// TwinCAT 3 PLC project Intecre_TwinSafeModels
// Title: Intecre.TwinSAFE.Models
// Company: Intecre Ltd
// Author: Mark Lazarides
// ProjectVersion: 0.5.0.3
// Description: Functional models of the TwinSAFE logic function blocks and TwinSAFE group, for trialling safety applications and their interaction with the standard PLC. 0.4.2.0 - T_SafeFunctionBlockBase sets State to Run / Stop before Process; user FBs need no State logic. 0.4.1.0 - corrects call issue with Example_UserFBs 0.4.0.0 - Adds the eight channel (EL1918) and two channel (EL2912) terminal models. 0.3.0.0 - Adds User FB examples, demonstrating extension.
// ProgramVersion: 3.1.4026.25
// libraries:
//   Intecre.Utilities, * (Intecre Ltd)
//   Tc2_Standard, * (Beckhoff Automation GmbH)
//   Tc2_System, * (Beckhoff Automation GmbH)
//   Tc3_Module, * (Beckhoff Automation GmbH)
//   TcUnit, * (www.tcunit.org)
// project tree:
//   / PlcTask.TcTTO
//   Core/ F_NormaliseSafeInput.TcPOU, F_SafeResetTimeOk.TcPOU, F_SafeInputValue.TcPOU, T_SafeConnection.TcPOU, T_SafeFunctionBlockBase.TcPOU, T_SafeGroup.TcPOU, T_SafeInputPair.TcPOU, T_SafeInputTerminal.TcPOU, T_SafeInputTerminal8.TcPOU, T_SafeOutputTerminal.TcPOU, T_SafeOutputTerminal2.TcPOU
//   DUTs/ E_SafeConnectionError.TcDUT, E_SafeConnectionState.TcDUT, E_SafeEdmState.TcDUT, E_SafeFbState.TcDUT, E_SafeGroupDiag.TcDUT, E_SafeGroupState.TcDUT, E_SafeLatchState.TcDUT, E_SafeMonState.TcDUT, E_SafeMutingState.TcDUT, E_SafeTonState.TcDUT, E_SafeTwoHandState.TcDUT, ST_SafeConnShutdownParameters.TcDUT, ST_SafeEStopParameters.TcDUT, ST_SafeEdmParameters.TcDUT, ST_SafeLatchParameters.TcDUT, ST_SafeLogicParameters.TcDUT, ST_SafeMonParameters.TcDUT, ST_SafeMutingParameters.TcDUT, ST_SafeOpModeParameters.TcDUT, ST_SafeTimerParameters.TcDUT, ST_SafeTwoHandParameters.TcDUT
//   Examples/Example_UserFbs/ T_SafePulse_UserFB.TcPOU, T_SafeRTrig_UserFB.TcPOU
//   Examples/ PRG_EStopExample.TcPOU, PRG_EStopExample_CFC.TcPOU
//   FunctionBlocks/ T_SafeAnd.TcPOU, T_SafeConnShutdown.TcPOU, T_SafeDecouple.TcPOU, T_SafeEStop.TcPOU, T_SafeEdm.TcPOU, T_SafeMon.TcPOU, T_SafeMuting.TcPOU, T_SafeOpMode.TcPOU, T_SafeOr.TcPOU, T_SafeRs.TcPOU, T_SafeSr.TcPOU, T_SafeTof.TcPOU, T_SafeTon.TcPOU, T_SafeTwoHand.TcPOU, T_SafeXor.TcPOU
//   Params/ SafeModelParams.TcGVL
//   Project Information/ F_GetCompany.TcPOU, F_GetTitle.TcPOU, F_GetVersion.TcPOU
//   Tests/ T_SafeCfcTestSuite.TcPOU, PRG_TestRunner.TcPOU, T_SafeAnd_Tests.TcPOU, T_SafeAnd_Tests_CFC.TcPOU, T_SafeConnShutdown_Tests.TcPOU, T_SafeConnShutdown_Tests_CFC.TcPOU, T_SafeConnection_Tests.TcPOU, T_SafeConnection_Tests_CFC.TcPOU, T_SafeDecouple_Tests.TcPOU, T_SafeDecouple_Tests_CFC.TcPOU, T_SafeEStop_Tests.TcPOU, T_SafeEStop_Tests_CFC.TcPOU, T_SafeEdm_Tests.TcPOU, T_SafeEdm_Tests_CFC.TcPOU, T_SafeGroup_Tests.TcPOU, T_SafeGroup_Tests_CFC.TcPOU, T_SafeInputPair_Tests.TcPOU, T_SafeInputPair_Tests_CFC.TcPOU, T_SafeInputTerminal8_Tests.TcPOU, T_SafeMon_Tests.TcPOU, T_SafeMon_Tests_CFC.TcPOU, T_SafeMuting_Tests.TcPOU, T_SafeMuting_Tests_CFC.TcPOU, T_SafeOpMode_Tests.TcPOU, T_SafeOpMode_Tests_CFC.TcPOU, T_SafeOr_Tests.TcPOU, T_SafeOr_Tests_CFC.TcPOU, T_SafeOutputTerminal2_Tests.TcPOU, T_SafeRs_Tests.TcPOU, T_SafeRs_Tests_CFC.TcPOU, T_SafeSr_Tests.TcPOU, T_SafeSr_Tests_CFC.TcPOU, T_SafeTof_Tests.TcPOU, T_SafeTof_Tests_CFC.TcPOU, T_SafeTon_Tests.TcPOU, T_SafeTon_Tests_CFC.TcPOU, T_SafeTwoHand_Tests.TcPOU, T_SafeTwoHand_Tests_CFC.TcPOU, T_SafeXor_Tests.TcPOU, T_SafeXor_Tests_CFC.TcPOU
//   Tests/User_FB_Tests/ T_SafePulse_UserFB_Tests.TcPOU, T_SafePulse_UserFB_Tests_CFC.TcPOU, T_SafeRTrig_UserFB_Tests.TcPOU, T_SafeRTrig_UserFB_Tests_CFC.TcPOU
//   Version/ Global_Version.TcGVL
// real-time tasks:
//   TASK PlcTask: cycle T#10ms, priority 20, ADS port 350

CONFIGURATION Intecre_TwinSafeModels
    RESOURCE PLC ON TwinCAT3
        TASK PlcTask(INTERVAL := T#10ms, PRIORITY := 20);
        PROGRAM PRG_TestRunner WITH PlcTask : PRG_TestRunner;
        PROGRAM PRG_EStopExample WITH PlcTask : PRG_EStopExample;
        PROGRAM PRG_EStopExample_CFC WITH PlcTask : PRG_EStopExample_CFC;
    END_RESOURCE
END_CONFIGURATION

// ---- DUTs/E_SafeConnectionError.TcDUT
// TwinSAFE connection error codes (low nibble of the connection Diag byte).
{attribute 'qualified_only'}
{attribute 'to_string'}
TYPE
E_SafeConnectionError :
(
    NoError := 0,
    InvalidCommand := 1,
    UnknownCommand := 2,
    InvalidConnectionId := 3,
    InvalidCrc := 4,
    WatchdogElapsed := 5,
    InvalidFsoeAddress := 6,
    InvalidData := 7,
    InvalidComParameterLength := 8,
    InvalidComParameters := 9,
    InvalidUserParameterLength := 10,
    InvalidUserParameters := 11,
    FsoeMasterReset := 12,
    SlaveModuleError := 13,
    OutputModuleError := 14,
    SlaveNotStarted := 15
) BYTE;
END_TYPE

// ---- DUTs/E_SafeConnectionState.TcDUT
// TwinSAFE (FSoE) connection state codes.
{attribute 'qualified_only'}
{attribute 'to_string'}
TYPE
E_SafeConnectionState :
(
    Reset := 100,
    Session := 101,
    Connection := 102,
    Parameter := 103,
    Data := 104,
    Shutdown := 105,
    ShutdownDeactive := 106
) BYTE;
END_TYPE

// ---- DUTs/E_SafeEdmState.TcDUT
// FB EDM state codes.
{attribute 'qualified_only'}
{attribute 'to_string'}
TYPE
E_SafeEdmState :
(
    Undefined := 0,
    Stop := 2,
    Error := 4,
    Reset := 5,
    MonOff := 14,
    MonOn := 15
) BYTE;
END_TYPE

// ---- DUTs/E_SafeFbState.TcDUT
// TwinSAFE function block state codes shared by most FBs (Map State value).
// Error is also the state of a block whose configuration the TwinSAFE Safety Editor refuses (too few
// inputs connected, a required input unwired, an invalid EDM reset time): the block then sets Error,
// diagnostic bit 15 (16#8000), which no TwinSAFE FB uses, and stays in Error through every ErrAck.
// See T_SafeFunctionBlockBase.
{attribute 'qualified_only'}
{attribute 'to_string'}
TYPE
E_SafeFbState :
(
    Undefined := 0,
    Run := 1,
    Stop := 2,
    Safe := 3,
    Error := 4,
    Reset := 5,
    Start := 6,
    ErrorDelay := 7,
    DelayOut := 8
) BYTE;
END_TYPE

// ---- DUTs/E_SafeGroupDiag.TcDUT
// TwinSAFE group diagnostic codes (EL/EJ6910).
{attribute 'qualified_only'}
{attribute 'to_string'}
TYPE
E_SafeGroupDiag :
(
    NoError := 0,
    FbError := 1,
    ComError := 2,
    ModuleError := 3,
    CmpError := 4,
    DeactivateError := 5,
    RestartError := 6
) BYTE;
END_TYPE

// ---- DUTs/E_SafeGroupState.TcDUT
// TwinSAFE group state codes (EL/EJ6910).
{attribute 'qualified_only'}
{attribute 'to_string'}
TYPE
E_SafeGroupState :
(
    Undefined := 0,
    Run := 1,
    Stop := 2,
    Safe := 3,
    Error := 4,
    Reset := 5,
    Start := 6,
    StopError := 7,
    Deactive := 16,
    WaitComError := 17
) BYTE;
END_TYPE

// ---- DUTs/E_SafeLatchState.TcDUT
// FB RS and FB SR state codes.
{attribute 'qualified_only'}
{attribute 'to_string'}
TYPE
E_SafeLatchState :
(
    Undefined := 0,
    Stop := 2,
    Safe := 3,
    Set := 9
) BYTE;
END_TYPE

// ---- DUTs/E_SafeMonState.TcDUT
// FB MON state codes.
{attribute 'qualified_only'}
{attribute 'to_string'}
TYPE
E_SafeMonState :
(
    Undefined := 0,
    Run := 1,
    Stop := 2,
    Safe := 3,
    Error := 4,
    Reset := 5,
    Start := 6,
    ErrorDelay := 7,
    DelayOut := 8,
    FuncTest := 9
) BYTE;
END_TYPE

// ---- DUTs/E_SafeMutingState.TcDUT
// FB MUTING state codes.
{attribute 'qualified_only'}
{attribute 'to_string'}
TYPE
E_SafeMutingState :
(
    Undefined := 0,
    Run := 1,
    Stop := 2,
    Safe := 3,
    Error := 4,
    Reset := 5,
    DelayOut := 8,
    Muting1 := 9,
    Muting2 := 10,
    Muting3 := 11,
    Muting4 := 12,
    Muting5 := 13,
    Muting6 := 14,
    Muting7 := 15,
    Muting8 := 16,
    Muting9 := 17
) BYTE;
END_TYPE

// ---- DUTs/E_SafeTonState.TcDUT
// FB TON state codes.
{attribute 'qualified_only'}
{attribute 'to_string'}
TYPE
E_SafeTonState :
(
    Undefined := 0,
    Run := 1,
    Stop := 2,
    Safe := 3,
    DelayIn := 9
) BYTE;
END_TYPE

// ---- DUTs/E_SafeTwoHandState.TcDUT
// FB TWOHAND state codes.
{attribute 'qualified_only'}
{attribute 'to_string'}
TYPE
E_SafeTwoHandState :
(
    Undefined := 0,
    Run := 1,
    Stop := 2,
    Safe := 3,
    Error := 4,
    Reset := 5,
    OneButton := 11,
    TwoButton := 12,
    Release := 13
) BYTE;
END_TYPE

// ---- DUTs/ST_SafeConnShutdownParameters.TcDUT
// Parameters of FB CONNECTION SHUTDOWN.
TYPE
ST_SafeConnShutdownParameters :
STRUCT
    Deactivate1MakeContact : BOOL;
    Deactivate2MakeContact : BOOL;
    DiscrepancyTime : TIME;
    SafeInputsAfterDiscError : BOOL; // Safety Editor checkbox 'Safe Inputs after Disc Error', FALSE for a new block:
        // TRUE makes both channels of the pair that raised a discrepancy error return to the safe state together
        // before ErrAck can clear it
END_STRUCT
END_TYPE

// ---- DUTs/ST_SafeEStopParameters.TcDUT
// Parameters of FB ESTOP (port and FB properties of the Safety Editor).
// Ports are active when connected; a pair is two channel when both ports are connected.
TYPE
ST_SafeEStopParameters :
STRUCT
    EStopIn1MakeContact : BOOL; // FALSE = break contact (0 requests the safe state); TRUE = make contact
    EStopIn2MakeContact : BOOL;
    EStopIn3MakeContact : BOOL;
    EStopIn4MakeContact : BOOL;
    EStopIn5MakeContact : BOOL;
    EStopIn6MakeContact : BOOL;
    EStopIn7MakeContact : BOOL;
    EStopIn8MakeContact : BOOL;
    DiscrepancyTime1 : TIME; // EStopIn1 / EStopIn2. T#0S = no discrepancy monitoring
    DiscrepancyTime2 : TIME; // EStopIn3 / EStopIn4
    DiscrepancyTime3 : TIME; // EStopIn5 / EStopIn6
    DiscrepancyTime4 : TIME; // EStopIn7 / EStopIn8
    DelayTime : TIME; // switch-off delay of EStopDelOut
    Edm1ResetTime : TIME; // EL6910: EDM1 must drop within this time of EStopOut switching on. T#0S disables
    Edm2ResetTime : TIME;
    SafeInputsAfterDiscError : BOOL; // Safety Editor checkbox, FALSE for a new block; the EL6910 always applies
        // 'Safe Inputs after Disc Error' to ESTOP whatever the box says (only the EL6900 honours it, and the editor
        // warns when it is TRUE under an EL6910), so the model ignores this value and always behaves as TRUE
END_STRUCT
END_TYPE

// ---- DUTs/ST_SafeEdmParameters.TcDUT
// Parameters of FB EDM.
TYPE
ST_SafeEdmParameters :
STRUCT
    Mon1MakeContact : BOOL;
    Mon2MakeContact : BOOL;
    SwitchOnTime : TIME; // Mon2 must become FALSE within this time of Mon1 rising. T#0S disables
    SwitchOffTime : TIME; // Mon2 must become TRUE within this time of Mon1 falling. T#0S disables
END_STRUCT
END_TYPE

// ---- DUTs/ST_SafeLatchParameters.TcDUT
// Parameters of FB RS and FB SR.
TYPE
ST_SafeLatchParameters :
STRUCT
    SetMakeContact : BOOL;
    ResetMakeContact : BOOL;
END_STRUCT
END_TYPE

// ---- DUTs/ST_SafeLogicParameters.TcDUT
// Parameters of FB AND and FB OR. Inputs are active when connected.
TYPE
ST_SafeLogicParameters :
STRUCT
    In1MakeContact : BOOL; // TRUE = the input is negated before the logic operation
    In2MakeContact : BOOL;
    In3MakeContact : BOOL;
    In4MakeContact : BOOL;
    In5MakeContact : BOOL;
    In6MakeContact : BOOL;
    In7MakeContact : BOOL;
    In8MakeContact : BOOL;
END_STRUCT
END_TYPE

// ---- DUTs/ST_SafeMonParameters.TcDUT
// Parameters of FB MON. Manual restart is active when the Restart port is connected.
TYPE
ST_SafeMonParameters :
STRUCT
    MonIn1MakeContact : BOOL;
    MonIn2MakeContact : BOOL;
    MonIn3MakeContact : BOOL;
    MonIn4MakeContact : BOOL;
    Secure1MakeContact : BOOL;
    Secure2MakeContact : BOOL;
    DiscrepancyTime1 : TIME; // MonIn1 / MonIn2
    DiscrepancyTime2 : TIME; // MonIn3 / MonIn4
    SecureDiscrepancyTime : TIME; // Secure1 / Secure2
    DelayTime : TIME; // switch-off delay of MonDelOut
    Edm1ResetTime : TIME;
    Edm2ResetTime : TIME;
    ManualFunctionTest : BOOL; // every connected MonIn pair must request the safe state once after start
    SafeInputsAfterDiscError : BOOL; // Safety Editor checkbox 'Safe Inputs after Disc Error', FALSE for a new block:
        // TRUE makes both channels of the pair that raised a discrepancy error return to the safe state together
        // before ErrAck can clear it
END_STRUCT
END_TYPE

// ---- DUTs/ST_SafeMutingParameters.TcDUT
// Parameters of FB MUTING.
TYPE
ST_SafeMutingParameters :
STRUCT
    SequentialInputs : BOOL; // TRUE: single-channel muting sensors in sequence; FALSE: two two-channel sensors
    MutingIn1MakeContact : BOOL;
    MutingIn2MakeContact : BOOL;
    MutingIn3MakeContact : BOOL;
    MutingIn4MakeContact : BOOL;
    OSSDIn1MakeContact : BOOL;
    OSSDIn2MakeContact : BOOL;
    MutingDiscrepancyTime1 : TIME; // MutingIn1 / MutingIn2 (parallel mode)
    MutingDiscrepancyTime2 : TIME; // MutingIn3 / MutingIn4 (parallel mode)
    OssdDiscrepancyTime : TIME; // OSSDIn1 / OSSDIn2
    FilterTime : TIME; // debounce of the muting inputs (max 500 ms)
    MaxMutingTime : TIME; // max duration of a muting sequence (max 10 min). T#0S disables
    DelayTime : TIME; // switch-off delay of MuteDelOut (max 30 s)
    Edm1ResetTime : TIME;
    Edm2ResetTime : TIME;
    BackwardsMode : BOOL; // EL6910: sequence may also run from the last sensor to the first
    OssdCheckOptional : BOOL; // EL6910: protective device is not part of the sequence check
    SafeInputsAfterDiscError : BOOL; // Safety Editor checkbox 'Safe Inputs after Disc Error', FALSE for a new block:
        // TRUE makes both channels of the pair that raised a discrepancy error return to the safe state together
        // before ErrAck can clear it
END_STRUCT
END_TYPE

// ---- DUTs/ST_SafeOpModeParameters.TcDUT
// Parameters of FB OPMODE. Manual restart is active when the Restart port is connected.
TYPE
ST_SafeOpModeParameters :
STRUCT
    DiscrepancyTime : TIME; // max time during a mode change with none or several inputs set. T#0S disables
END_STRUCT
END_TYPE

// ---- DUTs/ST_SafeTimerParameters.TcDUT
// Parameters of FB TON and FB TOF.
TYPE
ST_SafeTimerParameters :
STRUCT
    MakeContact : BOOL;
    DelayTime : TIME;
END_STRUCT
END_TYPE

// ---- DUTs/ST_SafeTwoHandParameters.TcDUT
// Parameters of FB TWOHAND.
TYPE
ST_SafeTwoHandParameters :
STRUCT
    Twohand1MakeContact : BOOL;
    Twohand2MakeContact : BOOL;
    Twohand3MakeContact : BOOL;
    Twohand4MakeContact : BOOL;
    DiscrepancyTime1 : TIME; // Twohand1 / Twohand2
    DiscrepancyTime2 : TIME; // Twohand3 / Twohand4
    HandDiscrepancyTime : TIME; // max time between actuation of the two hands (max 2500 ms). T#0S disables
    SafeInputsAfterDiscError : BOOL; // Safety Editor checkbox 'Safe Inputs after Disc Error', FALSE for a new block:
        // TRUE makes both channels of the pair that raised a discrepancy error return to the safe state together
        // before ErrAck can clear it
END_STRUCT
END_TYPE

// ---- Params/SafeModelParams.TcGVL
// Library parameters of Intecre.TwinSAFE.Models: the project-wide defaults, set per project in the
// Library Manager's parameter view without rebuilding the library. A parameter list must be constant,
// so the run-time switch lives on T_SafeGroup (RaiseOnRefusedConfiguration), initialised from here.
{attribute 'qualified_only'}
VAR_GLOBAL CONSTANT
    // Default of T_SafeGroup.RaiseOnRefusedConfiguration for every group. TRUE: a block of the group whose
    // configuration the TwinSAFE Safety Editor refuses (see T_SafeFunctionBlockBase) raises
    // RTSEXCPT_IO_CONFIG_ERROR with F_RaiseException after it has reported Error, so the controller stops
    // on the first cycle unless the call is in a __TRY block. FALSE: the block only reports Error,
    // State = Error and diagnostic bit 15, and logs the fault once.
    RAISE_ON_REFUSED_CONFIGURATION : BOOL := FALSE;
END_VAR

// ---- Version/Global_Version.TcGVL
{attribute 'TcGenerated'}
{attribute 'no-analysis'}
{attribute 'linkalways'}
// This function has been automatically generated from the project information.
VAR_GLOBAL CONSTANT
	{attribute 'const_non_replaced'}
	stLibVersion_Intecre_TwinSAFE_Models : ST_LibVersion := (iMajor := 0, iMinor := 5, iBuild := 0, iRevision := 3, nFlags := 0, sVersion := '0.5.0.3');
END_VAR

// ---- Tests/PRG_TestRunner.TcPOU
// Runs every TcUnit test suite in the library.
PROGRAM PRG_TestRunner
VAR
    safeAndTests                    : T_SafeAnd_Tests;
    safeInputPairTests              : T_SafeInputPair_Tests;
    safeOrTests                     : T_SafeOr_Tests;
    safeXorTests                    : T_SafeXor_Tests;
    safeDecoupleTests               : T_SafeDecouple_Tests;
    safeOpModeTests                 : T_SafeOpMode_Tests;
    safeRsTests                     : T_SafeRs_Tests;
    safeSrTests                     : T_SafeSr_Tests;
    safeTonTests                    : T_SafeTon_Tests;
    safeTofTests                    : T_SafeTof_Tests;
    safeEdmTests                    : T_SafeEdm_Tests;
    safeEStopTests                  : T_SafeEStop_Tests;
    safeMonTests                    : T_SafeMon_Tests;
    safeTwoHandTests                : T_SafeTwoHand_Tests;
    safeMutingTests                 : T_SafeMuting_Tests;
    safeConnectionTests             : T_SafeConnection_Tests;
    safeInputTerminal8Tests         : T_SafeInputTerminal8_Tests;
    safeOutputTerminal2Tests        : T_SafeOutputTerminal2_Tests;
    safeConnShutdownTests           : T_SafeConnShutdown_Tests;
    safeGroupTests                  : T_SafeGroup_Tests;
    safePulseUserFbTests            : T_SafePulse_UserFB_Tests;
    safeRTrigUserFbTests            : T_SafeRTrig_UserFB_Tests;

    // CFC twins of the suites above
    safeAndTestsCfc                 : T_SafeAnd_Tests_CFC;
    safeInputPairTestsCfc           : T_SafeInputPair_Tests_CFC;
    safeOrTestsCfc                  : T_SafeOr_Tests_CFC;
    safeXorTestsCfc                 : T_SafeXor_Tests_CFC;
    safeDecoupleTestsCfc            : T_SafeDecouple_Tests_CFC;
    safeOpModeTestsCfc              : T_SafeOpMode_Tests_CFC;
    safeRsTestsCfc                  : T_SafeRs_Tests_CFC;
    safeSrTestsCfc                  : T_SafeSr_Tests_CFC;
    safeTonTestsCfc                 : T_SafeTon_Tests_CFC;
    safeTofTestsCfc                 : T_SafeTof_Tests_CFC;
    safeEdmTestsCfc                 : T_SafeEdm_Tests_CFC;
    safeEStopTestsCfc               : T_SafeEStop_Tests_CFC;
    safeMonTestsCfc                 : T_SafeMon_Tests_CFC;
    safeTwoHandTestsCfc             : T_SafeTwoHand_Tests_CFC;
    safeMutingTestsCfc              : T_SafeMuting_Tests_CFC;
    safeConnectionTestsCfc          : T_SafeConnection_Tests_CFC;
    safeConnShutdownTestsCfc        : T_SafeConnShutdown_Tests_CFC;
    safeGroupTestsCfc               : T_SafeGroup_Tests_CFC;
    safePulseUserFbTestsCfc         : T_SafePulse_UserFB_Tests_CFC;
    safeRTrigUserFbTestsCfc         : T_SafeRTrig_UserFB_Tests_CFC;
END_VAR

// Intecre.Utilities logs nothing until a project sets LogConfig.LogLevel; Error lets the
// refused-configuration lines of the configuration tests through to the TwinCAT log.
LogConfig.LogLevel := E_LogSeverity.Error;
TcUnit.RUN();

END_PROGRAM

// ---- Tests/T_SafeAnd_Tests.TcPOU
FUNCTION_BLOCK T_SafeAnd_Tests EXTENDS TcUnit.FB_TestSuite
VAR
    // Test_AllConnectedInputsTrueGivesRun
    group_1 : T_SafeGroup;
    fb_1 : T_SafeAnd(group := group_1);
    // Test_OneInputFalseGivesSafe
    group_2 : T_SafeGroup;
    fb_2 : T_SafeAnd(group := group_2);
    // Test_UnconnectedInputsIgnoredAndMakeContactNegated
    group_3 : T_SafeGroup;
    fb_3 : T_SafeAnd(group := group_3) := (Parameters := (In2MakeContact := TRUE));
    // Test_StoppedGivesNoOutput
    group_4 : T_SafeGroup;
    fb_4 : T_SafeAnd(group := group_4);
    // Test_OneConnectedInputIsRefused
    group_5 : T_SafeGroup;
    fb_5 : T_SafeAnd(group := group_5);
    // Test_RaiseOnRefusedConfigurationStopsHard
    group_6 : T_SafeGroup;
    fb_6 : T_SafeAnd(group := group_6);
END_VAR

Test_AllConnectedInputsTrueGivesRun();
Test_OneInputFalseGivesSafe();
Test_UnconnectedInputsIgnoredAndMakeContactNegated();
Test_StoppedGivesNoOutput();
Test_OneConnectedInputIsRefused();
Test_RaiseOnRefusedConfigurationStopsHard();

METHOD PRIVATE Test_AllConnectedInputsTrueGivesRun
TcUnit.TEST(__POUNAME());
// act
group_1(Run := TRUE);
fb_1(AndIn1 := TRUE, AndIn2 := TRUE);
// assert
AssertEquals_BOOL(Expected := TRUE, Actual := fb_1.AndOut, Message := 'output on when all connected inputs are 1');
AssertEquals_BYTE(Expected := TO_BYTE(E_SafeFbState.Run), Actual := fb_1.State, Message := 'state RUN');
TEST_FINISHED_NAMED(__POUNAME());
END_METHOD

METHOD PRIVATE Test_OneInputFalseGivesSafe
TcUnit.TEST(__POUNAME());
// act
group_2(Run := TRUE);
fb_2(AndIn1 := TRUE, AndIn2 := FALSE);
// assert
AssertEquals_BOOL(Expected := FALSE, Actual := fb_2.AndOut, Message := 'output off when a connected input is 0');
AssertEquals_BYTE(Expected := TO_BYTE(E_SafeFbState.Safe), Actual := fb_2.State, Message := 'state SAFE');
TEST_FINISHED_NAMED(__POUNAME());
END_METHOD

METHOD PRIVATE Test_StoppedGivesNoOutput
TcUnit.TEST(__POUNAME());
// act
group_4(Run := FALSE);
fb_4(AndIn1 := TRUE, AndIn2 := TRUE);
// assert
AssertEquals_BOOL(Expected := FALSE, Actual := fb_4.AndOut, Message := 'no output while the group is stopped');
AssertEquals_BYTE(Expected := TO_BYTE(E_SafeFbState.Stop), Actual := fb_4.State, Message := 'state STOP');
TEST_FINISHED_NAMED(__POUNAME());
END_METHOD

METHOD PRIVATE Test_UnconnectedInputsIgnoredAndMakeContactNegated
TcUnit.TEST(__POUNAME());
// act: AndIn3..8 unconnected, AndIn2 make contact at 0 (released)
group_3(Run := TRUE);
fb_3(AndIn1 := TRUE, AndIn2 := FALSE);
// assert
AssertEquals_BOOL(Expected := TRUE, Actual := fb_3.AndOut, Message := 'unconnected inputs ignored, make contact negated');
TEST_FINISHED_NAMED(__POUNAME());
END_METHOD

METHOD PRIVATE Test_OneConnectedInputIsRefused
TcUnit.TEST(__POUNAME());
// arrange / act: AndIn1 is the only connected input, which the Safety Editor refuses
group_5(Run := TRUE);
fb_5(AndIn1 := TRUE);
group_5(Run := TRUE);
fb_5(AndIn1 := TRUE);
// assert
AssertEquals_BOOL(Expected := TRUE, Actual := fb_5.Error, Message := 'configuration error reported');
AssertEquals_BYTE(Expected := TO_BYTE(E_SafeFbState.Error), Actual := fb_5.State, Message := 'state ERROR');
AssertEquals_WORD(Expected := WORD#16#8000, Actual := fb_5.Diag, Message := 'diag bit 15 configuration refused');
AssertEquals_BOOL(Expected := FALSE, Actual := fb_5.AndOut, Message := 'AndOut stays at its safe value');
AssertEquals_BOOL(Expected := TRUE, Actual := group_5.FbErr, Message := 'the group sees an FB error');
// act: ErrAck 0 -> 1 -> 0 does not clear a configuration error
group_5(Run := TRUE, ErrAck := TRUE);
fb_5(AndIn1 := TRUE);
group_5(Run := TRUE, ErrAck := TRUE);
fb_5(AndIn1 := TRUE);
group_5(Run := TRUE, ErrAck := FALSE);
fb_5(AndIn1 := TRUE);
AssertEquals_BOOL(Expected := TRUE, Actual := fb_5.Error, Message := 'error not acknowledged');
AssertEquals_WORD(Expected := WORD#16#8000, Actual := fb_5.Diag, Message := 'diag bit 15 kept');
TEST_FINISHED_NAMED(__POUNAME());
END_METHOD

METHOD PRIVATE Test_RaiseOnRefusedConfigurationStopsHard
VAR
    exc : __SYSTEM.ExceptionCode;
    caught : __SYSTEM.ExceptionCode;
END_VAR
TcUnit.TEST(__POUNAME());
// arrange: a one-input AND, the group's opt-in hard stop switched on for this call only
caught := __SYSTEM.ExceptionCode.RTSEXCPT_NOEXCEPTION;
group_6.RaiseOnRefusedConfiguration := TRUE;
// act
__TRY
    group_6(Run := TRUE);
    fb_6(AndIn1 := TRUE);
__CATCH(exc)
    caught := exc;
__FINALLY
    group_6.RaiseOnRefusedConfiguration := FALSE;
__ENDTRY
// assert: the code given to F_RaiseException does not reach __CATCH on TwinCAT 3.1 4026 (the x64
// usermode runtime delivered 16#E8940001 instead of RTSEXCPT_IO_CONFIG_ERROR), so only the arrival
// of an exception is checked; the block's own outputs carry the reason
AssertEquals_BOOL(Expected := TRUE, Actual := (caught <> __SYSTEM.ExceptionCode.RTSEXCPT_NOEXCEPTION), Message := 'an exception was raised and caught');
AssertEquals_BOOL(Expected := TRUE, Actual := fb_6.Error, Message := 'error reported before the exception');
AssertEquals_BYTE(Expected := TO_BYTE(E_SafeFbState.Error), Actual := fb_6.State, Message := 'state ERROR');
AssertEquals_WORD(Expected := WORD#16#8000, Actual := fb_6.Diag, Message := 'diag bit 15 configuration refused');
TEST_FINISHED_NAMED(__POUNAME());
END_METHOD

END_FUNCTION_BLOCK

// ---- Core/T_SafeGroup.TcPOU
// Model of a TwinSAFE group (EL/EJ6910 semantics).
// Function blocks and connections join the group at construction (FB_init group reference) and the
// group reads their outputs, so nothing needs wiring beyond the standard PLC signals.
// Call the group before its members each cycle. Declare the group before its members.
// RaiseOnRefusedConfiguration (default SafeModelParams.RAISE_ON_REFUSED_CONFIGURATION) makes a member
// whose configuration the Safety Editor refuses stop the controller with F_RaiseException after it has
// reported Error; see T_SafeFunctionBlockBase.
FUNCTION_BLOCK T_SafeGroup
VAR_INPUT
    Run : BOOL := TRUE; // Run/Stop. Link to a standard PLC variable.
    ErrAck : BOOL; // Error acknowledge (FALSE -> TRUE -> FALSE). Link to a standard PLC variable.
    ModuleFault : BOOL; // error input from another module (e.g. EK1960)
END_VAR
VAR_OUTPUT
    ComErr : BOOL; // communication error in at least one connection
    FbErr : BOOL; // at least one FB is in the ERROR state
    OutErr : BOOL; // not used (local outputs only exist on KL6904)
    OtherErr : BOOL; // ModuleFault
    ComStartup : BOOL; // at least one connection is starting up
    FbDeactive : BOOL; // group deactivated by customising (not modelled, always FALSE)
    FbRun : BOOL; // all FBs are in the RUN state
    InRun : BOOL; // the group is in the RUN state (FbRun of the members)
    State : BYTE; // group state code (Map State)
    Diag : BYTE; // group diagnostic code (Map Diag)
    RegistrationRefused : BOOL; // a block or connection could not join because the group is full (MAX_FUNCTION_BLOCKS, MAX_CONNECTIONS): the model is then incomplete, never expected in use
END_VAR
VAR CONSTANT
    MAX_FUNCTION_BLOCKS : UINT := 256;
    MAX_CONNECTIONS : UINT := 64;
END_VAR
VAR
    _functionBlocks : ARRAY[1..MAX_FUNCTION_BLOCKS] OF POINTER TO T_SafeFunctionBlockBase;
    _functionBlockCount : UINT;
    _connections : ARRAY[1..MAX_CONNECTIONS] OF POINTER TO T_SafeConnection;
    _connectionCount : UINT;
    _state : E_SafeGroupState := E_SafeGroupState.Stop;
    _prevState : E_SafeGroupState;
    _errAckPrev : BOOL;
    _errAckFallingEdge : BOOL;
    _anyFbError : BOOL;
    _allFbsRunning : BOOL;
    _anyComError : BOOL;
    _anyComStartup : BOOL;
    _anyError : BOOL;
    _raiseOnRefusedConfiguration : BOOL := SafeModelParams.RAISE_ON_REFUSED_CONFIGURATION;
END_VAR

_errAckFallingEdge := NOT ErrAck AND _errAckPrev;
_errAckPrev        := ErrAck;
ScanMembers();
_anyError := _anyFbError OR _anyComError OR ModuleFault;

CASE _state OF
    E_SafeGroupState.Undefined,
    E_SafeGroupState.Stop:
        StateChanged();

        IF _anyError THEN
            _state := E_SafeGroupState.StopError;
        ELSIF Run THEN
            _state := SEL(_anyComStartup, E_SafeGroupState.Run, E_SafeGroupState.Start);
        END_IF

    E_SafeGroupState.StopError:
        StateChanged();

        IF Run THEN
            _state := E_SafeGroupState.Error;
        ELSIF NOT _anyError THEN
            _state := E_SafeGroupState.Stop;
        END_IF

    E_SafeGroupState.Start:
        StateChanged();

        IF _anyError THEN
            _state := E_SafeGroupState.Error;
        ELSIF NOT Run THEN
            _state := E_SafeGroupState.Stop;
        ELSIF NOT _anyComStartup THEN
            _state := E_SafeGroupState.Run;
        END_IF

    E_SafeGroupState.Run:
        StateChanged();

        IF _anyError THEN
            _state := E_SafeGroupState.Error;
        ELSIF NOT Run THEN
            _state := E_SafeGroupState.Stop;
        ELSIF _anyComStartup THEN
            _state := E_SafeGroupState.Start;
        END_IF

    E_SafeGroupState.Error:
        StateChanged();

        IF NOT Run THEN
            _state := E_SafeGroupState.StopError;
        ELSIF ErrAck AND NOT _anyError THEN
            _state := E_SafeGroupState.Reset;
        END_IF

    E_SafeGroupState.Reset:
        StateChanged();

        IF _anyError THEN
            _state := E_SafeGroupState.Error;
        ELSIF _errAckFallingEdge THEN
            IF NOT Run THEN
                _state := E_SafeGroupState.Stop;
            ELSIF _anyComStartup THEN
                _state := E_SafeGroupState.Start;
            ELSE
                _state := E_SafeGroupState.Run;
            END_IF
        END_IF

ELSE
    _state := E_SafeGroupState.Stop;
END_CASE

ComErr     := _anyComError;
FbErr      := _anyFbError;
OutErr     := FALSE;
OtherErr   := ModuleFault;
ComStartup := _anyComStartup;
FbDeactive := FALSE;
FbRun      := _allFbsRunning;
InRun      := (_state = E_SafeGroupState.Run);
State      := TO_BYTE(_state);

IF _anyFbError THEN
    Diag := TO_BYTE(E_SafeGroupDiag.FbError);
ELSIF _anyComError THEN
    Diag := TO_BYTE(E_SafeGroupDiag.ComError);
ELSIF ModuleFault THEN
    Diag := TO_BYTE(E_SafeGroupDiag.ModuleError);
ELSE
    Diag := TO_BYTE(E_SafeGroupDiag.NoError);
END_IF

PROPERTY ConnectionCount : UINT
GET
ConnectionCount := _connectionCount;
END_GET
END_PROPERTY

PROPERTY FunctionBlockCount : UINT
GET
FunctionBlockCount := _functionBlockCount;
END_GET
END_PROPERTY

PROPERTY GroupState : E_SafeGroupState
GET
GroupState := _state;
END_GET
END_PROPERTY

// TRUE: a member whose configuration the TwinSAFE Safety Editor refuses raises RTSEXCPT_IO_CONFIG_ERROR
// (F_RaiseException) after reporting Error, so the controller stops unless the call is in a __TRY block.
// Starts at SafeModelParams.RAISE_ON_REFUSED_CONFIGURATION; set it per group from project code or a test.
PROPERTY RaiseOnRefusedConfiguration : BOOL
GET
RaiseOnRefusedConfiguration := _raiseOnRefusedConfiguration;
END_GET
SET
_raiseOnRefusedConfiguration := RaiseOnRefusedConfiguration;
END_SET
END_PROPERTY

// Called by T_SafeConnection.FB_init. Not part of the public interface.
METHOD INTERNAL RegisterConnection
VAR_INPUT
    connection : REFERENCE TO T_SafeConnection;
END_VAR
VAR
    i : UINT;
END_VAR
FOR i := 1 TO _connectionCount DO
    IF _connections[i] = ADR(connection) THEN
        RETURN;
    END_IF
END_FOR

IF _connectionCount >= MAX_CONNECTIONS THEN
    RegistrationRefused := TRUE;
    RETURN;
END_IF

_connectionCount               := _connectionCount + 1;
_connections[_connectionCount] := ADR(connection);
END_METHOD

// Called by T_SafeFunctionBlockBase.FB_init. Not part of the public interface.
METHOD INTERNAL RegisterFunctionBlock
VAR_INPUT
    functionBlock : REFERENCE TO T_SafeFunctionBlockBase;
END_VAR
VAR
    i : UINT;
END_VAR
FOR i := 1 TO _functionBlockCount DO
    IF _functionBlocks[i] = ADR(functionBlock) THEN
        RETURN;
    END_IF
END_FOR

IF _functionBlockCount >= MAX_FUNCTION_BLOCKS THEN
    RegistrationRefused := TRUE;
    RETURN;
END_IF

_functionBlockCount                  := _functionBlockCount + 1;
_functionBlocks[_functionBlockCount] := ADR(functionBlock);
END_METHOD

// Reads the outputs of the registered function blocks and connections.
METHOD PRIVATE ScanMembers
VAR
    i : UINT;
END_VAR
_anyFbError    := FALSE;
_allFbsRunning := (_functionBlockCount > 0);

FOR i := 1 TO _functionBlockCount DO
    _anyFbError    := _anyFbError OR _functionBlocks[i]^.Error;
    _allFbsRunning := _allFbsRunning AND _functionBlocks[i]^.IsRunning;
END_FOR

_anyComError   := FALSE;
_anyComStartup := FALSE;

FOR i := 1 TO _connectionCount DO
    _anyComError   := _anyComError OR _connections[i]^.ComError;
    _anyComStartup := _anyComStartup OR _connections[i]^.InStartup;
END_FOR
END_METHOD

METHOD PRIVATE StateChanged : BOOL
IF _prevState = _state THEN
    RETURN;
END_IF

_prevState   := _state;
StateChanged := TRUE;
END_METHOD

END_FUNCTION_BLOCK

// ---- Core/T_SafeFunctionBlockBase.TcPOU
// Common behaviour of every modelled TwinSAFE function block.
// A block belongs to a TwinSAFE group from construction: declare it as
//     eStop : T_SafeEStop(group := safetyGroup);
// It registers with the group, takes FbRun (group in RUN) and ErrAck from it, and the group
// reads its Error and IsRunning outputs. Declare the group before its members.
// Derived classes implement Process(). Before Process() the base sets State to Run while the group
// runs and to Stop otherwise, so a block built only from other blocks needs no State logic; a block
// with states of its own overwrites State in Process(), and writes Error and Diag when it has them.
//
// Configuration check. The Safety Editor refuses some wirings and parameter values at project verify
// (an AND with one input, an SR with Reset unwired, an EDM reset time that is not a multiple of 10 ms).
// A block with such a rule overrides ConfigurationOk() and writes the editor's message to
// _configurationFault when the rule is broken. The base then runs the block as a stopped block (outputs
// at their safe value), reports Error with State = Error and diagnostic bit 15 (16#8000, a bit no
// TwinSAFE FB uses), logs the fault once through the Intecre.Utilities logger with the instance name in
// front (taken from the private T_NamedBase member _log; the project has to set LogConfig.LogLevel to
// Error or lower, as the logger is silent by default), and keeps the error through every ErrAck: a
// configuration error cannot be acknowledged away, only rewired.
// With the group's RaiseOnRefusedConfiguration TRUE (default SafeModelParams.RAISE_ON_REFUSED_CONFIGURATION,
// a library parameter) the base also raises RTSEXCPT_IO_CONFIG_ERROR with F_RaiseException after
// reporting, so a simulation stops hard on the first cycle unless the call sits in a __TRY block
// (a __CATCH on 4026 receives a TwinCAT code, not RTSEXCPT_IO_CONFIG_ERROR; check Error and Diag).
FUNCTION_BLOCK ABSTRACT T_SafeFunctionBlockBase
VAR_OUTPUT
    Error : BOOL; // FB Error output
    State : BYTE; // FB state code (Map State)
    Diag : WORD; // FB diagnostic bits (Map Diag)
    IsRunning : BOOL; // FB in the RUN state
END_VAR
VAR CONSTANT
    CONFIGURATION_REFUSED_DIAG_BIT : INT := 15; // Diag bit set while the Safety Editor would refuse the configuration
END_VAR
VAR
    _group : REFERENCE TO T_SafeGroup;
    _fbRun : BOOL; // group in RUN
    _errAck : BOOL; // group error acknowledge
    _errAckPrev : BOOL;
    _errAckRisingEdge : BOOL;
    _errAckFallingEdge : BOOL;
    _configurationRefused : BOOL; // ConfigurationOk() returned FALSE this cycle
    _configurationFault : T_MaxString; // the editor's message for the broken rule, written by ConfigurationOk()
    _configurationLogged : BOOL; // the fault has been logged (once per instance)
    _log : T_NamedBase; // supplies the instance path for the log line; its InstanceName ends in ._log, which ReportRefusedConfiguration trims
END_VAR

IF __ISVALIDREF(_group) THEN
    _fbRun  := _group.InRun;
    _errAck := _group.ErrAck;
ELSE
    // not (yet) in a group: behaves as a stopped block until SetGroupReference is called
    _fbRun  := FALSE;
    _errAck := FALSE;
END_IF

_configurationRefused := NOT ConfigurationOk();

IF _configurationRefused THEN
    // the Safety Editor refuses this wiring or parameter set: the block runs as a stopped block, so its
    // outputs take their safe value, and the error reported below is not acknowledged
    _fbRun  := FALSE;
    _errAck := FALSE;
END_IF

_errAckRisingEdge  := _errAck AND NOT _errAckPrev;
_errAckFallingEdge := NOT _errAck AND _errAckPrev;
_errAckPrev        := _errAck;
// default state: Run while the group runs, else Stop. Blocks with states of their own overwrite it in
// Process(). Error and Diag are not reset here: they latch until ErrAck in TwinSAFE, so only the block
// that raised them clears them.
State := TO_BYTE(SEL(_fbRun, E_SafeFbState.Stop, E_SafeFbState.Run));
Process();

IF _configurationRefused THEN
    Error := TRUE;
    State := TO_BYTE(E_SafeFbState.Error);
    SetDiagBit(CONFIGURATION_REFUSED_DIAG_BIT);
END_IF

IsRunning := (State = TO_BYTE(E_SafeFbState.Run));

IF _configurationRefused THEN
    ReportRefusedConfiguration();
END_IF

METHOD PROTECTED ClearDiagBit
VAR_INPUT
    bitIndex : INT;
END_VAR
Diag := Diag AND NOT SHL(WORD#1, bitIndex);
END_METHOD

// TRUE when the block is wired and parameterised as the TwinSAFE Safety Editor accepts it. A block
// with a rule overrides this method; when the rule is broken it writes the editor's own message to
// _configurationFault and returns FALSE. The base then reports the block in Error (see the header).
METHOD PROTECTED ConfigurationOk : BOOL
ConfigurationOk := TRUE;
END_METHOD

METHOD FB_init : BOOL
VAR_INPUT
    bInitRetains : BOOL;
    bInCopyCode : BOOL;
    group : REFERENCE TO T_SafeGroup; // the TwinSAFE group this block belongs to
END_VAR
SetGroupReference(
    bInCopyCode := bInCopyCode,
    group := group
);
END_METHOD

METHOD PROTECTED ABSTRACT Process
END_METHOD

// Logs the refused configuration once per instance as '<instance>: <block type>: <editor's rule> (...)',
// the instance being _log.InstanceName minus its own '._log' segment, then stops the controller with
// RTSEXCPT_IO_CONFIG_ERROR when the group's RaiseOnRefusedConfiguration asks for it (a block without a
// group follows the library parameter). Called after Error, State and Diag have been written, so a
// __CATCH sees the block already in Error. The logger is Intecre.Utilities' F_LogError, which is silent
// until the project sets LogConfig.LogLevel.
METHOD PRIVATE ReportRefusedConfiguration
VAR
    instance : T_MaxString;
    raise : BOOL;
END_VAR
VAR CONSTANT
    MEMBER_SUFFIX : STRING := '._log';
END_VAR
IF NOT _configurationLogged THEN
    _configurationLogged := TRUE;
    instance := _log.InstanceName;

    IF RIGHT(instance, LEN(MEMBER_SUFFIX)) = MEMBER_SUFFIX THEN
        instance := LEFT(instance, LEN(instance) - LEN(MEMBER_SUFFIX));
    END_IF

    F_LogError(CONCAT(CONCAT(instance, ': '), CONCAT(_configurationFault, ' (the TwinSAFE Safety Editor refuses this configuration)')));
END_IF

IF __ISVALIDREF(_group) THEN
    raise := _group.RaiseOnRefusedConfiguration;
ELSE
    raise := SafeModelParams.RAISE_ON_REFUSED_CONFIGURATION;
END_IF

IF raise THEN
    F_RaiseException(TO_UDINT(__SYSTEM.ExceptionCode.RTSEXCPT_IO_CONFIG_ERROR));
END_IF
END_METHOD

METHOD PROTECTED SetDiagBit
VAR_INPUT
    bitIndex : INT;
END_VAR
Diag := Diag OR SHL(WORD#1, bitIndex);
END_METHOD

// Assigns the block to a TwinSAFE group and registers it there. Called by FB_init; call it
// yourself from the FB_init of a composite (user) block to pass its group on to the blocks it
// contains, which were declared with the composite's own _group before that reference was valid.
// Registering twice with the same group is harmless. Returns TRUE when the group was valid.
METHOD PUBLIC SetGroupReference : BOOL
VAR_INPUT
    bInCopyCode : BOOL;
    group : REFERENCE TO T_SafeGroup; // the TwinSAFE group this block belongs to
END_VAR
IF NOT __ISVALIDREF(group) THEN
    RETURN;
END_IF

_group REF= group;

IF NOT bInCopyCode THEN
    group.RegisterFunctionBlock(THIS^);
END_IF

SetGroupReference := TRUE;
END_METHOD

END_FUNCTION_BLOCK

// ---- Core/T_SafeConnection.TcPOU
// Simulated TwinSAFE (FSoE) connection between the logic and a safe I/O terminal or another logic.
// Belongs to a group from construction:  conn : T_SafeConnection(group := safetyGroup);
// Starts up through Reset -> Session -> Connection -> Parameter -> Data once the group runs.
// Communication errors are injected with InjectComError and cleared by the group ErrAck
// (plus ComErrAck when ComErrAckActive is set).
FUNCTION_BLOCK T_SafeConnection
VAR_INPUT
    ComErrAck : BOOL; // connection specific acknowledgement (EL6910 option ComErrAckActive)
    LocalShutdown : BOOL; // shutdown requested by FB CONNECTION SHUTDOWN (set through its reference)
    PartnerShutdown : BOOL; // simulates a shutdown command received from the FSoE partner
    InjectComError : BOOL; // rising edge simulates an FSoE communication error
    InjectErrorCode : E_SafeConnectionError := E_SafeConnectionError.WatchdogElapsed;
    StartupTime : TIME := T#300MS; // simulated time from Reset to Data
    ComErrAckActive : BOOL; // connection needs its own ComErrAck in addition to the group ErrAck
END_VAR
VAR_OUTPUT
    ComError : BOOL;
    InStartup : BOOL;
    InDataState : BOOL;
    OutputsEnabled : BOOL; // in the Data state with the group in RUN: the only time a safe output terminal passes its SafeOut values (a group in STOP or ERROR switches every output of the group off)
    IsShutdown : BOOL;
    State : BYTE; // connection state code 100..106
    Diag : BYTE; // connection diagnostic byte
END_VAR
VAR
    _group : REFERENCE TO T_SafeGroup;
    _state : E_SafeConnectionState := E_SafeConnectionState.Reset;
    _prevState : E_SafeConnectionState;
    _errorCode : E_SafeConnectionError;
    _groupAcknowledged : BOOL;
    _comErrAcked : BOOL;
    _errAckPrev : BOOL;
    _comErrAckPrev : BOOL;
    _injectPrev : BOOL;
    _startupTimer : TON;
END_VAR

IF NOT __ISVALIDREF(_group) THEN
    RETURN; // not (yet) assigned to a group: stays in its initial (fail-safe) state
END_IF

IF _group.ErrAck AND NOT _errAckPrev THEN
    _groupAcknowledged := TRUE;
END_IF

_errAckPrev := _group.ErrAck;

IF ComErrAck AND NOT _comErrAckPrev THEN
    _comErrAcked := TRUE;
END_IF

_comErrAckPrev := ComErrAck;

IF InjectComError AND NOT _injectPrev THEN
    ComError           := TRUE;
    _errorCode         := InjectErrorCode;
    _groupAcknowledged := FALSE;
    _comErrAcked       := FALSE;
    _state             := E_SafeConnectionState.Reset;
END_IF

_injectPrev := InjectComError;

// A communication error is cleared once the group (and if required the connection) has acknowledged.
IF ComError AND _groupAcknowledged AND (NOT ComErrAckActive OR _comErrAcked) THEN
    ComError           := FALSE;
    _errorCode         := E_SafeConnectionError.NoError;
    _groupAcknowledged := FALSE;
    _comErrAcked       := FALSE;
END_IF

RunStateMachine();

InStartup := NOT ComError
                 AND (_state = E_SafeConnectionState.Reset
                 OR _state = E_SafeConnectionState.Session
                 OR _state = E_SafeConnectionState.Connection
                 OR _state = E_SafeConnectionState.Parameter);

InDataState := (_state = E_SafeConnectionState.Data);
OutputsEnabled := InDataState AND _group.InRun;
IsShutdown  := (_state = E_SafeConnectionState.Shutdown) OR (_state = E_SafeConnectionState.ShutdownDeactive);
State       := TO_BYTE(_state);
Diag        := TO_BYTE(_errorCode);

IF InStartup THEN
    Diag := Diag OR 16#40;
END_IF

IF ComError THEN
    Diag := Diag OR 16#10;
END_IF

METHOD FB_init : BOOL
VAR_INPUT
    bInitRetains : BOOL;
    bInCopyCode : BOOL;
    group : REFERENCE TO T_SafeGroup; // the TwinSAFE group this connection is assigned to
END_VAR
SetGroupReference(
    bInCopyCode := bInCopyCode,
    group := group
);
END_METHOD

// Assigns the connection to a TwinSAFE group and registers it there. Called by FB_init; call it
// yourself from the FB_init of a composite (user) block to pass its group on to a connection it
// contains, which was declared with the composite's own _group before that reference was valid.
// Registering twice with the same group is harmless. Returns TRUE when the group was valid.
METHOD PUBLIC SetGroupReference : BOOL
VAR_INPUT
    bInCopyCode : BOOL;
    group : REFERENCE TO T_SafeGroup; // the TwinSAFE group this connection is assigned to
END_VAR
IF NOT __ISVALIDREF(group) THEN
    RETURN;
END_IF

_group REF= group;

IF NOT bInCopyCode THEN
    group.RegisterConnection(THIS^);
END_IF

SetGroupReference := TRUE;
END_METHOD

METHOD PRIVATE RunStateMachine
VAR
    stepTime : TIME;
END_VAR
stepTime := UDINT_TO_TIME(TIME_TO_UDINT(StartupTime) / 3);

CASE _state OF
    E_SafeConnectionState.Reset:
        IF StateChanged() THEN
            _startupTimer(IN := FALSE, PT := stepTime);
        END_IF

        IF _group.Run AND NOT ComError THEN
            _state := E_SafeConnectionState.Session;
        END_IF

    E_SafeConnectionState.Session:
        IF StateChanged() THEN
            _startupTimer(IN := FALSE, PT := stepTime);
        END_IF

        _startupTimer(IN := TRUE, PT := stepTime);

        IF _startupTimer.Q THEN
            _state := E_SafeConnectionState.Connection;
        END_IF

    E_SafeConnectionState.Connection:
        IF StateChanged() THEN
            _startupTimer(IN := FALSE, PT := stepTime);
        END_IF

        _startupTimer(IN := TRUE, PT := stepTime);

        IF _startupTimer.Q THEN
            _state := E_SafeConnectionState.Parameter;
        END_IF

    E_SafeConnectionState.Parameter:
        IF StateChanged() THEN
            _startupTimer(IN := FALSE, PT := stepTime);
        END_IF

        _startupTimer(IN := TRUE, PT := stepTime);

        IF _startupTimer.Q THEN
            _state := E_SafeConnectionState.Data;
        END_IF

    E_SafeConnectionState.Data:
        StateChanged();

        IF LocalShutdown THEN
            _state := E_SafeConnectionState.ShutdownDeactive;
        ELSIF PartnerShutdown THEN
            _state := E_SafeConnectionState.Shutdown;
        END_IF

    E_SafeConnectionState.Shutdown:
        StateChanged();

        IF NOT PartnerShutdown THEN
            _state := E_SafeConnectionState.Reset;
        END_IF

    E_SafeConnectionState.ShutdownDeactive:
        StateChanged();

        IF NOT LocalShutdown THEN
            _state := E_SafeConnectionState.Reset;
        END_IF
END_CASE
END_METHOD

METHOD PRIVATE StateChanged : BOOL
IF _prevState = _state THEN
    RETURN;
END_IF

_prevState   := _state;
StateChanged := TRUE;
END_METHOD

END_FUNCTION_BLOCK

// ---- FunctionBlocks/T_SafeAnd.TcPOU
// Model of the TwinSAFE FB AND. Connected inputs are active; AndIn1 may be a standard PLC signal.
// The Safety Editor refuses an AND with fewer than two AndIn ports connected: the model then reports
// Error with diagnostic bit 15 instead of running (see T_SafeFunctionBlockBase).
{attribute 'reflection'}
FUNCTION_BLOCK T_SafeAnd EXTENDS T_SafeFunctionBlockBase
VAR_INPUT
    AndIn1 : BOOL;
    AndIn2 : BOOL;
    AndIn3 : BOOL;
    AndIn4 : BOOL;
    AndIn5 : BOOL;
    AndIn6 : BOOL;
    AndIn7 : BOOL;
    AndIn8 : BOOL;
    Parameters : ST_SafeLogicParameters;
END_VAR
VAR_OUTPUT
    AndOut : BOOL;
END_VAR
VAR
    {attribute 'is_connected' := 'AndIn1'}
    _andIn1Connected : BOOL;
    {attribute 'is_connected' := 'AndIn2'}
    _andIn2Connected : BOOL;
    {attribute 'is_connected' := 'AndIn3'}
    _andIn3Connected : BOOL;
    {attribute 'is_connected' := 'AndIn4'}
    _andIn4Connected : BOOL;
    {attribute 'is_connected' := 'AndIn5'}
    _andIn5Connected : BOOL;
    {attribute 'is_connected' := 'AndIn6'}
    _andIn6Connected : BOOL;
    {attribute 'is_connected' := 'AndIn7'}
    _andIn7Connected : BOOL;
    {attribute 'is_connected' := 'AndIn8'}
    _andIn8Connected : BOOL;
    _state : E_SafeFbState := E_SafeFbState.Stop;
END_VAR

SUPER^();

// At least two AndIn ports must be connected (Safety Editor: "AND does not have at least 2 input ports active and connected").
METHOD PROTECTED ConfigurationOk : BOOL
VAR
    connectedInputs : USINT;
END_VAR
connectedInputs := BOOL_TO_USINT(_andIn1Connected)
    + BOOL_TO_USINT(_andIn2Connected)
    + BOOL_TO_USINT(_andIn3Connected)
    + BOOL_TO_USINT(_andIn4Connected)
    + BOOL_TO_USINT(_andIn5Connected)
    + BOOL_TO_USINT(_andIn6Connected)
    + BOOL_TO_USINT(_andIn7Connected)
    + BOOL_TO_USINT(_andIn8Connected);

IF connectedInputs < 2 THEN
    _configurationFault := 'T_SafeAnd: AND does not have at least 2 input ports active and connected';
    RETURN;
END_IF

ConfigurationOk := TRUE;
END_METHOD

METHOD PROTECTED Process
VAR
    result : BOOL;
END_VAR
result := TRUE;
result := result AND F_NormaliseSafeInput(_andIn1Connected, Parameters.In1MakeContact, AndIn1);
result := result AND F_NormaliseSafeInput(_andIn2Connected, Parameters.In2MakeContact, AndIn2);
result := result AND F_NormaliseSafeInput(_andIn3Connected, Parameters.In3MakeContact, AndIn3);
result := result AND F_NormaliseSafeInput(_andIn4Connected, Parameters.In4MakeContact, AndIn4);
result := result AND F_NormaliseSafeInput(_andIn5Connected, Parameters.In5MakeContact, AndIn5);
result := result AND F_NormaliseSafeInput(_andIn6Connected, Parameters.In6MakeContact, AndIn6);
result := result AND F_NormaliseSafeInput(_andIn7Connected, Parameters.In7MakeContact, AndIn7);
result := result AND F_NormaliseSafeInput(_andIn8Connected, Parameters.In8MakeContact, AndIn8);

IF NOT _fbRun THEN
    _state := E_SafeFbState.Stop;
ELSIF result THEN
    _state := E_SafeFbState.Run;
ELSE
    _state := E_SafeFbState.Safe;
END_IF

AndOut := (_state = E_SafeFbState.Run);
Error  := FALSE;
Diag   := 0;
State  := TO_BYTE(_state);
END_METHOD

END_FUNCTION_BLOCK

// ---- Core/F_NormaliseSafeInput.TcPOU
// Applies the port configuration to a raw input value.
// Result TRUE means "not requesting the safe state" (the released / healthy condition).
// An unconnected (inactive) port never requests the safe state.
FUNCTION F_NormaliseSafeInput : BOOL
VAR_INPUT
    active : BOOL; // port is connected
    makeContact : BOOL; // FALSE = break contact (0 requests the safe state), TRUE = make contact (signal negated)
    value : BOOL;
END_VAR

IF NOT active THEN
    F_NormaliseSafeInput := TRUE;
    RETURN;
END_IF

F_NormaliseSafeInput := value XOR makeContact;

END_FUNCTION

// ---- Tests/T_SafeInputPair_Tests.TcPOU
FUNCTION_BLOCK T_SafeInputPair_Tests EXTENDS TcUnit.FB_TestSuite
VAR
    // Test_DiscrepancyErrorAfterTimeoutAndResetAfterSafeInputs
    pair_5 : T_SafeInputPair;
    state_5 : INT := 10;
    waitTimer_5 : TON;
END_VAR

Test_InactivePairNeverRequestsSafeState();
Test_BreakContactRequestsSafeStateOnZero();
Test_MakeContactRequestsSafeStateOnOne();
Test_TwoChannelRequestsSafeStateIfEitherChannelLow();
Test_DiscrepancyErrorAfterTimeoutAndResetAfterSafeInputs();

METHOD PRIVATE Test_BreakContactRequestsSafeStateOnZero
VAR
    pair : T_SafeInputPair;
END_VAR
TcUnit.TEST(__POUNAME());
// act
pair(In1 := FALSE, Active1 := TRUE, Monitor := TRUE);
// assert
AssertEquals_BOOL(Expected := TRUE, Actual := pair.SafeStateRequested, Message := 'break contact at 0 must request the safe state');
pair(In1 := TRUE, Active1 := TRUE, Monitor := TRUE);
AssertEquals_BOOL(Expected := FALSE, Actual := pair.SafeStateRequested, Message := 'break contact at 1 must not request the safe state');
TEST_FINISHED_NAMED(__POUNAME());
END_METHOD

METHOD PRIVATE Test_DiscrepancyErrorAfterTimeoutAndResetAfterSafeInputs
TcUnit.TEST(__POUNAME());
waitTimer_5();

CASE state_5 OF
    10:
        // arrange
        state_5 := 20;
        waitTimer_5(IN := TRUE, PT := T#50MS);
    20:
        // act: channels disagree for less than the discrepancy time
        pair_5(
            In1 := TRUE,
            In2 := FALSE,
            Active1 := TRUE,
            Active2 := TRUE,
            Monitor := TRUE,
            SafeInputsAfterDiscError := TRUE,
            DiscrepancyTime := T#100MS
        );

        IF NOT waitTimer_5.Q THEN
            RETURN;
        END_IF

        waitTimer_5(IN := FALSE);
        // assert
        AssertEquals_BOOL(Expected := FALSE, Actual := pair_5.DiscrepancyError, Message := 'no error before the discrepancy time');
        state_5 := 30;
        waitTimer_5(IN := TRUE, PT := T#200MS);
    30:
        pair_5(
            In1 := TRUE,
            In2 := FALSE,
            Active1 := TRUE,
            Active2 := TRUE,
            Monitor := TRUE,
            SafeInputsAfterDiscError := TRUE,
            DiscrepancyTime := T#100MS
        );

        IF NOT waitTimer_5.Q THEN
            RETURN;
        END_IF

        waitTimer_5(IN := FALSE);
        // assert
        AssertEquals_BOOL(Expected := TRUE, Actual := pair_5.DiscrepancyError, Message := 'error after the discrepancy time');
        AssertEquals_BOOL(Expected := TRUE, Actual := pair_5.AwaitingSafeInputs, Message := 'error waits for both channels safe');
        // act: acknowledge while a channel is still high
        pair_5(
            In1 := TRUE,
            In2 := FALSE,
            Active1 := TRUE,
            Active2 := TRUE,
            Monitor := TRUE,
            SafeInputsAfterDiscError := TRUE,
            DiscrepancyTime := T#100MS,
            Acknowledge := TRUE
        );

        AssertEquals_BOOL(Expected := TRUE, Actual := pair_5.DiscrepancyError, Message := 'acknowledge refused while a channel is still high');
        // act: both channels safe, then acknowledge
        pair_5(
            In1 := FALSE,
            In2 := FALSE,
            Active1 := TRUE,
            Active2 := TRUE,
            Monitor := TRUE,
            SafeInputsAfterDiscError := TRUE,
            DiscrepancyTime := T#100MS,
            Acknowledge := TRUE
        );

        AssertEquals_BOOL(Expected := FALSE, Actual := pair_5.DiscrepancyError, Message := 'error cleared once both channels were safe');
        TEST_FINISHED_NAMED(__POUNAME());
        state_5 := 10;
END_CASE
END_METHOD

METHOD PRIVATE Test_InactivePairNeverRequestsSafeState
VAR
    pair : T_SafeInputPair;
END_VAR
TcUnit.TEST(__POUNAME());
// act
pair(In1 := FALSE, In2 := FALSE, Active1 := FALSE, Active2 := FALSE, Monitor := TRUE);
// assert
AssertEquals_BOOL(Expected := FALSE, Actual := pair.SafeStateRequested, Message := 'inactive pair must not request the safe state');
AssertEquals_BOOL(Expected := FALSE, Actual := pair.IsActive, Message := 'pair should be inactive');
TEST_FINISHED_NAMED(__POUNAME());
END_METHOD

METHOD PRIVATE Test_MakeContactRequestsSafeStateOnOne
VAR
    pair : T_SafeInputPair;
END_VAR
TcUnit.TEST(__POUNAME());
// act
pair(In1 := TRUE, Active1 := TRUE, MakeContact1 := TRUE, Monitor := TRUE);
// assert
AssertEquals_BOOL(Expected := TRUE, Actual := pair.SafeStateRequested, Message := 'make contact at 1 must request the safe state');
TEST_FINISHED_NAMED(__POUNAME());
END_METHOD

METHOD PRIVATE Test_TwoChannelRequestsSafeStateIfEitherChannelLow
VAR
    pair : T_SafeInputPair;
END_VAR
TcUnit.TEST(__POUNAME());
// act
pair(
    In1 := TRUE,
    In2 := FALSE,
    Active1 := TRUE,
    Active2 := TRUE,
    Monitor := TRUE,
    SafeInputsAfterDiscError := TRUE
);

// assert
AssertEquals_BOOL(Expected := TRUE, Actual := pair.SafeStateRequested, Message := 'one low channel must request the safe state');
AssertEquals_BOOL(Expected := FALSE, Actual := pair.DiscrepancyError, Message := 'no discrepancy monitoring without a discrepancy time');
pair(
    In1 := TRUE,
    In2 := TRUE,
    Active1 := TRUE,
    Active2 := TRUE,
    Monitor := TRUE,
    SafeInputsAfterDiscError := TRUE
);

AssertEquals_BOOL(Expected := FALSE, Actual := pair.SafeStateRequested, Message := 'both channels high must not request the safe state');
TEST_FINISHED_NAMED(__POUNAME());
END_METHOD

END_FUNCTION_BLOCK

// ---- Core/T_SafeInputPair.TcPOU
// Evaluates a one- or two-channel FB input pair with optional discrepancy monitoring,
// exactly as the TwinSAFE FBs treat their paired inputs (EStopIn1/2, MonIn1/2, Twohand1/2 ...).
// Internal helper used by the modelled FBs.
FUNCTION_BLOCK T_SafeInputPair
VAR_INPUT
    In1 : BOOL;
    In2 : BOOL;
    Active1 : BOOL; // channel 1 port is connected
    Active2 : BOOL; // channel 2 port is connected
    MakeContact1 : BOOL;
    MakeContact2 : BOOL;
    DiscrepancyTime : TIME; // T#0S = two channel without discrepancy monitoring
    Monitor : BOOL; // discrepancy monitoring runs only while TRUE (FB executed by a running group)
    SafeInputsAfterDiscError : BOOL; // both channels must be safe together before a discrepancy error can be acknowledged
    Acknowledge : BOOL; // clear a discrepancy error this cycle if permitted
END_VAR
VAR_OUTPUT
    Channel1 : BOOL; // normalised: TRUE = not requesting the safe state
    Channel2 : BOOL;
    IsActive : BOOL;
    IsTwoChannel : BOOL;
    AllTrue : BOOL; // all active channels TRUE (TRUE when inactive)
    AllFalse : BOOL; // all active channels FALSE (FALSE when inactive)
    SafeStateRequested : BOOL;
    DiscrepancyError : BOOL;
    AwaitingSafeInputs : BOOL;
END_VAR
VAR
    _discrepancyTimer : TON;
END_VAR

Channel1     := F_NormaliseSafeInput(Active1, MakeContact1, In1);
Channel2     := F_NormaliseSafeInput(Active2, MakeContact2, In2);
IsActive     := Active1 OR Active2;
IsTwoChannel := Active1 AND Active2;

IF Monitor AND IsTwoChannel AND DiscrepancyTime > T#0S THEN
    _discrepancyTimer(IN := (Channel1 <> Channel2), PT := DiscrepancyTime);

    IF _discrepancyTimer.Q AND NOT DiscrepancyError THEN
        DiscrepancyError   := TRUE;
        AwaitingSafeInputs := SafeInputsAfterDiscError;
    END_IF
ELSE
    _discrepancyTimer(IN := FALSE, PT := DiscrepancyTime);
END_IF

IF AwaitingSafeInputs AND NOT Channel1 AND NOT Channel2 THEN
    AwaitingSafeInputs := FALSE;
END_IF

IF Acknowledge AND DiscrepancyError AND NOT AwaitingSafeInputs THEN
    DiscrepancyError := FALSE;
    _discrepancyTimer(IN := FALSE, PT := DiscrepancyTime);
END_IF

AllTrue            := Channel1 AND Channel2;
AllFalse           := IsActive AND (NOT Active1 OR NOT Channel1) AND (NOT Active2 OR NOT Channel2);
SafeStateRequested := NOT AllTrue;

END_FUNCTION_BLOCK

// ---- Tests/T_SafeOr_Tests.TcPOU
FUNCTION_BLOCK T_SafeOr_Tests EXTENDS TcUnit.FB_TestSuite
VAR
    // Test_AnyConnectedInputTrueGivesRun
    group_1 : T_SafeGroup;
    fb_1 : T_SafeOr(group := group_1);
    // Test_AllFalseGivesSafe
    group_2 : T_SafeGroup;
    fb_2 : T_SafeOr(group := group_2);
    // Test_OneConnectedInputIsRefused
    group_3 : T_SafeGroup;
    fb_3 : T_SafeOr(group := group_3);
END_VAR

Test_AnyConnectedInputTrueGivesRun();
Test_AllFalseGivesSafe();
Test_OneConnectedInputIsRefused();

METHOD PRIVATE Test_AllFalseGivesSafe
TcUnit.TEST(__POUNAME());
// act
group_2(Run := TRUE);
fb_2(OrIn1 := FALSE, OrIn2 := FALSE);
// assert
AssertEquals_BOOL(Expected := FALSE, Actual := fb_2.OrOut, Message := 'output off when all connected inputs are 0');
AssertEquals_BYTE(Expected := TO_BYTE(E_SafeFbState.Safe), Actual := fb_2.State, Message := 'state SAFE');
TEST_FINISHED_NAMED(__POUNAME());
END_METHOD

METHOD PRIVATE Test_AnyConnectedInputTrueGivesRun
TcUnit.TEST(__POUNAME());
// act
group_1(Run := TRUE);
fb_1(OrIn1 := FALSE, OrIn2 := TRUE);
// assert
AssertEquals_BOOL(Expected := TRUE, Actual := fb_1.OrOut, Message := 'output on when any connected input is 1');
TEST_FINISHED_NAMED(__POUNAME());
END_METHOD

METHOD PRIVATE Test_OneConnectedInputIsRefused
TcUnit.TEST(__POUNAME());
// arrange / act: OrIn1 is the only connected input, which the Safety Editor refuses
group_3(Run := TRUE);
fb_3(OrIn1 := TRUE);
group_3(Run := TRUE);
fb_3(OrIn1 := TRUE);
// assert
AssertEquals_BOOL(Expected := TRUE, Actual := fb_3.Error, Message := 'configuration error reported');
AssertEquals_BYTE(Expected := TO_BYTE(E_SafeFbState.Error), Actual := fb_3.State, Message := 'state ERROR');
AssertEquals_WORD(Expected := WORD#16#8000, Actual := fb_3.Diag, Message := 'diag bit 15 configuration refused');
AssertEquals_BOOL(Expected := FALSE, Actual := fb_3.OrOut, Message := 'OrOut stays at its safe value');
AssertEquals_BOOL(Expected := TRUE, Actual := group_3.FbErr, Message := 'the group sees an FB error');
// act: ErrAck 0 -> 1 -> 0 does not clear a configuration error
group_3(Run := TRUE, ErrAck := TRUE);
fb_3(OrIn1 := TRUE);
group_3(Run := TRUE, ErrAck := TRUE);
fb_3(OrIn1 := TRUE);
group_3(Run := TRUE, ErrAck := FALSE);
fb_3(OrIn1 := TRUE);
AssertEquals_BOOL(Expected := TRUE, Actual := fb_3.Error, Message := 'error not acknowledged');
AssertEquals_WORD(Expected := WORD#16#8000, Actual := fb_3.Diag, Message := 'diag bit 15 kept');
TEST_FINISHED_NAMED(__POUNAME());
END_METHOD

END_FUNCTION_BLOCK

// ---- FunctionBlocks/T_SafeOr.TcPOU
// Model of the TwinSAFE FB OR. Connected inputs are active.
// The Safety Editor refuses an OR with fewer than two OrIn ports connected: the model then reports
// Error with diagnostic bit 15 instead of running (see T_SafeFunctionBlockBase).
{attribute 'reflection'}
FUNCTION_BLOCK T_SafeOr EXTENDS T_SafeFunctionBlockBase
VAR_INPUT
    OrIn1 : BOOL;
    OrIn2 : BOOL;
    OrIn3 : BOOL;
    OrIn4 : BOOL;
    OrIn5 : BOOL;
    OrIn6 : BOOL;
    OrIn7 : BOOL;
    OrIn8 : BOOL;
    Parameters : ST_SafeLogicParameters;
END_VAR
VAR_OUTPUT
    OrOut : BOOL;
END_VAR
VAR
    {attribute 'is_connected' := 'OrIn1'}
    _orIn1Connected : BOOL;
    {attribute 'is_connected' := 'OrIn2'}
    _orIn2Connected : BOOL;
    {attribute 'is_connected' := 'OrIn3'}
    _orIn3Connected : BOOL;
    {attribute 'is_connected' := 'OrIn4'}
    _orIn4Connected : BOOL;
    {attribute 'is_connected' := 'OrIn5'}
    _orIn5Connected : BOOL;
    {attribute 'is_connected' := 'OrIn6'}
    _orIn6Connected : BOOL;
    {attribute 'is_connected' := 'OrIn7'}
    _orIn7Connected : BOOL;
    {attribute 'is_connected' := 'OrIn8'}
    _orIn8Connected : BOOL;
    _state : E_SafeFbState := E_SafeFbState.Stop;
END_VAR

SUPER^();

// At least two OrIn ports must be connected (Safety Editor: "OR does not have at least 2 input ports active and connected").
METHOD PROTECTED ConfigurationOk : BOOL
VAR
    connectedInputs : USINT;
END_VAR
connectedInputs := BOOL_TO_USINT(_orIn1Connected)
    + BOOL_TO_USINT(_orIn2Connected)
    + BOOL_TO_USINT(_orIn3Connected)
    + BOOL_TO_USINT(_orIn4Connected)
    + BOOL_TO_USINT(_orIn5Connected)
    + BOOL_TO_USINT(_orIn6Connected)
    + BOOL_TO_USINT(_orIn7Connected)
    + BOOL_TO_USINT(_orIn8Connected);

IF connectedInputs < 2 THEN
    _configurationFault := 'T_SafeOr: OR does not have at least 2 input ports active and connected';
    RETURN;
END_IF

ConfigurationOk := TRUE;
END_METHOD

METHOD PROTECTED Process
VAR
    result : BOOL;
END_VAR
result := FALSE;
result := result OR F_SafeInputValue(_orIn1Connected, Parameters.In1MakeContact, OrIn1);
result := result OR F_SafeInputValue(_orIn2Connected, Parameters.In2MakeContact, OrIn2);
result := result OR F_SafeInputValue(_orIn3Connected, Parameters.In3MakeContact, OrIn3);
result := result OR F_SafeInputValue(_orIn4Connected, Parameters.In4MakeContact, OrIn4);
result := result OR F_SafeInputValue(_orIn5Connected, Parameters.In5MakeContact, OrIn5);
result := result OR F_SafeInputValue(_orIn6Connected, Parameters.In6MakeContact, OrIn6);
result := result OR F_SafeInputValue(_orIn7Connected, Parameters.In7MakeContact, OrIn7);
result := result OR F_SafeInputValue(_orIn8Connected, Parameters.In8MakeContact, OrIn8);

IF NOT _fbRun THEN
    _state := E_SafeFbState.Stop;
ELSIF result THEN
    _state := E_SafeFbState.Run;
ELSE
    _state := E_SafeFbState.Safe;
END_IF

OrOut := (_state = E_SafeFbState.Run);
Error := FALSE;
Diag  := 0;
State := TO_BYTE(_state);
END_METHOD

END_FUNCTION_BLOCK

// ---- Core/F_SafeInputValue.TcPOU
// Applies the port configuration to a raw input value for ports that assert a function
// (Set, Reset, TonIn, OrIn, muting sensors ...). An unconnected port reads FALSE.
FUNCTION F_SafeInputValue : BOOL
VAR_INPUT
    active : BOOL;
    makeContact : BOOL;
    value : BOOL;
END_VAR

IF NOT active THEN
    F_SafeInputValue := FALSE;
    RETURN;
END_IF

F_SafeInputValue := value XOR makeContact;

END_FUNCTION

// ---- Tests/T_SafeXor_Tests.TcPOU
FUNCTION_BLOCK T_SafeXor_Tests EXTENDS TcUnit.FB_TestSuite
VAR
    // Test_ConnectedPairsAreExclusiveOr
    group_1 : T_SafeGroup;
    fb_1 : T_SafeXor(group := group_1);
END_VAR

Test_ConnectedPairsAreExclusiveOr();

METHOD PRIVATE Test_ConnectedPairsAreExclusiveOr
TcUnit.TEST(__POUNAME());
// act
group_1(Run := TRUE);
fb_1(Xor1In1 := TRUE, Xor2In1 := FALSE);
// assert
AssertEquals_BOOL(Expected := TRUE, Actual := fb_1.XorOut1, Message := 'connected pair 1 XOR');
AssertEquals_BOOL(Expected := FALSE, Actual := fb_1.XorOut2, Message := 'unconnected pair stays 0');
fb_1(Xor1In1 := TRUE, Xor2In1 := TRUE);
AssertEquals_BOOL(Expected := FALSE, Actual := fb_1.XorOut1, Message := 'both inputs 1 gives 0');
TEST_FINISHED_NAMED(__POUNAME());
END_METHOD

END_FUNCTION_BLOCK

// ---- FunctionBlocks/T_SafeXor.TcPOU
// Model of the TwinSAFE FB XOR: eight independent exclusive-or pairs. A pair is active when connected.
{attribute 'reflection'}
FUNCTION_BLOCK T_SafeXor EXTENDS T_SafeFunctionBlockBase
VAR_INPUT
    Xor1In1 : BOOL;
    Xor2In1 : BOOL;
    Xor1In2 : BOOL;
    Xor2In2 : BOOL;
    Xor1In3 : BOOL;
    Xor2In3 : BOOL;
    Xor1In4 : BOOL;
    Xor2In4 : BOOL;
    Xor1In5 : BOOL;
    Xor2In5 : BOOL;
    Xor1In6 : BOOL;
    Xor2In6 : BOOL;
    Xor1In7 : BOOL;
    Xor2In7 : BOOL;
    Xor1In8 : BOOL;
    Xor2In8 : BOOL;
END_VAR
VAR_OUTPUT
    XorOut1 : BOOL;
    XorOut2 : BOOL;
    XorOut3 : BOOL;
    XorOut4 : BOOL;
    XorOut5 : BOOL;
    XorOut6 : BOOL;
    XorOut7 : BOOL;
    XorOut8 : BOOL;
END_VAR
VAR
    {attribute 'is_connected' := 'Xor1In1'}
    _xor1In1Connected : BOOL;
    {attribute 'is_connected' := 'Xor1In2'}
    _xor1In2Connected : BOOL;
    {attribute 'is_connected' := 'Xor1In3'}
    _xor1In3Connected : BOOL;
    {attribute 'is_connected' := 'Xor1In4'}
    _xor1In4Connected : BOOL;
    {attribute 'is_connected' := 'Xor1In5'}
    _xor1In5Connected : BOOL;
    {attribute 'is_connected' := 'Xor1In6'}
    _xor1In6Connected : BOOL;
    {attribute 'is_connected' := 'Xor1In7'}
    _xor1In7Connected : BOOL;
    {attribute 'is_connected' := 'Xor1In8'}
    _xor1In8Connected : BOOL;
    {attribute 'is_connected' := 'Xor2In1'}
    _xor2In1Connected : BOOL;
    {attribute 'is_connected' := 'Xor2In2'}
    _xor2In2Connected : BOOL;
    {attribute 'is_connected' := 'Xor2In3'}
    _xor2In3Connected : BOOL;
    {attribute 'is_connected' := 'Xor2In4'}
    _xor2In4Connected : BOOL;
    {attribute 'is_connected' := 'Xor2In5'}
    _xor2In5Connected : BOOL;
    {attribute 'is_connected' := 'Xor2In6'}
    _xor2In6Connected : BOOL;
    {attribute 'is_connected' := 'Xor2In7'}
    _xor2In7Connected : BOOL;
    {attribute 'is_connected' := 'Xor2In8'}
    _xor2In8Connected : BOOL;
    _state : E_SafeFbState := E_SafeFbState.Stop;
END_VAR

SUPER^();

METHOD PROTECTED Process
VAR
    run : BOOL;
END_VAR
run     := _fbRun;
_state  := SEL(run, E_SafeFbState.Stop, E_SafeFbState.Run);
XorOut1 := run AND (_xor1In1Connected OR _xor2In1Connected) AND (Xor1In1 XOR Xor2In1);
XorOut2 := run AND (_xor1In2Connected OR _xor2In2Connected) AND (Xor1In2 XOR Xor2In2);
XorOut3 := run AND (_xor1In3Connected OR _xor2In3Connected) AND (Xor1In3 XOR Xor2In3);
XorOut4 := run AND (_xor1In4Connected OR _xor2In4Connected) AND (Xor1In4 XOR Xor2In4);
XorOut5 := run AND (_xor1In5Connected OR _xor2In5Connected) AND (Xor1In5 XOR Xor2In5);
XorOut6 := run AND (_xor1In6Connected OR _xor2In6Connected) AND (Xor1In6 XOR Xor2In6);
XorOut7 := run AND (_xor1In7Connected OR _xor2In7Connected) AND (Xor1In7 XOR Xor2In7);
XorOut8 := run AND (_xor1In8Connected OR _xor2In8Connected) AND (Xor1In8 XOR Xor2In8);
Error   := FALSE;
Diag    := 0;
State   := TO_BYTE(_state);
END_METHOD

END_FUNCTION_BLOCK

// ---- Tests/T_SafeDecouple_Tests.TcPOU
FUNCTION_BLOCK T_SafeDecouple_Tests EXTENDS TcUnit.FB_TestSuite
VAR
    // Test_InputsLoopedToOutputsOnlyWhenRunning
    group_1 : T_SafeGroup;
    fb_1 : T_SafeDecouple(group := group_1);
END_VAR

Test_InputsLoopedToOutputsOnlyWhenRunning();

METHOD PRIVATE Test_InputsLoopedToOutputsOnlyWhenRunning
TcUnit.TEST(__POUNAME());
// act
group_1(Run := TRUE);
fb_1(DecIn3 := TRUE);
// assert
AssertEquals_BOOL(Expected := TRUE, Actual := fb_1.DecOut3, Message := 'input looped to output');
group_1(Run := FALSE);
fb_1(DecIn3 := TRUE);
AssertEquals_BOOL(Expected := FALSE, Actual := fb_1.DecOut3, Message := 'output off while the group is stopped');
TEST_FINISHED_NAMED(__POUNAME());
END_METHOD

END_FUNCTION_BLOCK

// ---- FunctionBlocks/T_SafeDecouple.TcPOU
// Model of the TwinSAFE FB DECOUPLE: eight inputs looped one-to-one to eight outputs.
FUNCTION_BLOCK T_SafeDecouple EXTENDS T_SafeFunctionBlockBase
VAR_INPUT
    DecIn1 : BOOL;
    DecIn2 : BOOL;
    DecIn3 : BOOL;
    DecIn4 : BOOL;
    DecIn5 : BOOL;
    DecIn6 : BOOL;
    DecIn7 : BOOL;
    DecIn8 : BOOL;
END_VAR
VAR_OUTPUT
    DecOut1 : BOOL;
    DecOut2 : BOOL;
    DecOut3 : BOOL;
    DecOut4 : BOOL;
    DecOut5 : BOOL;
    DecOut6 : BOOL;
    DecOut7 : BOOL;
    DecOut8 : BOOL;
END_VAR
VAR
    _state : E_SafeFbState := E_SafeFbState.Stop;
END_VAR

SUPER^();

METHOD PROTECTED Process
VAR
    run : BOOL;
END_VAR
run     := _fbRun;
_state  := SEL(run, E_SafeFbState.Stop, E_SafeFbState.Run);
DecOut1 := run AND DecIn1;
DecOut2 := run AND DecIn2;
DecOut3 := run AND DecIn3;
DecOut4 := run AND DecIn4;
DecOut5 := run AND DecIn5;
DecOut6 := run AND DecIn6;
DecOut7 := run AND DecIn7;
DecOut8 := run AND DecIn8;
Error   := FALSE;
Diag    := 0;
State   := TO_BYTE(_state);
END_METHOD

END_FUNCTION_BLOCK

// ---- Tests/T_SafeOpMode_Tests.TcPOU
FUNCTION_BLOCK T_SafeOpMode_Tests EXTENDS TcUnit.FB_TestSuite
VAR
    // Test_ExactlyOneInputSelectsOutput
    group_1 : T_SafeGroup;
    fb_1 : T_SafeOpMode(group := group_1);
    // Test_ConnectedRestartRequiresRestartSequence
    group_2 : T_SafeGroup;
    fb_2 : T_SafeOpMode(group := group_2);
    // Test_SlowModeChangeGivesDiscrepancyError
    group_3 : T_SafeGroup;
    fb_3 : T_SafeOpMode(group := group_3) := (Parameters := (DiscrepancyTime := T#100MS));
    state_3 : INT := 10;
    waitTimer_3 : TON;
    // Test_OneConnectedInputIsRefused
    group_4 : T_SafeGroup;
    fb_4 : T_SafeOpMode(group := group_4);
END_VAR

Test_ExactlyOneInputSelectsOutput();
Test_ConnectedRestartRequiresRestartSequence();
Test_SlowModeChangeGivesDiscrepancyError();
Test_OneConnectedInputIsRefused();

METHOD PRIVATE Test_ConnectedRestartRequiresRestartSequence
TcUnit.TEST(__POUNAME());
// act
group_2(Run := TRUE);
fb_2(Restart := FALSE, OpIn1 := TRUE, OpIn2 := FALSE);
group_2(Run := TRUE);
fb_2(Restart := FALSE, OpIn1 := TRUE, OpIn2 := FALSE);
// assert
AssertEquals_BOOL(Expected := FALSE, Actual := fb_2.OpOut1, Message := 'no output before restart');
group_2(Run := TRUE);
fb_2(Restart := TRUE, OpIn1 := TRUE, OpIn2 := FALSE);
AssertEquals_BYTE(Expected := TO_BYTE(E_SafeFbState.Start), Actual := fb_2.State, Message := 'state START while restart held');
group_2(Run := TRUE);
fb_2(Restart := FALSE, OpIn1 := TRUE, OpIn2 := FALSE);
AssertEquals_BOOL(Expected := TRUE, Actual := fb_2.OpOut1, Message := 'output on after restart falling edge');
TEST_FINISHED_NAMED(__POUNAME());
END_METHOD

METHOD PRIVATE Test_ExactlyOneInputSelectsOutput
TcUnit.TEST(__POUNAME());
// act: STOP -> SAFE -> RUN (no Restart connected: automatic)
group_1(Run := TRUE);
fb_1(OpIn1 := FALSE, OpIn2 := TRUE);
group_1(Run := TRUE);
fb_1(OpIn1 := FALSE, OpIn2 := TRUE);
// assert
AssertEquals_BOOL(Expected := TRUE, Actual := fb_1.OpOut2, Message := 'selected mode output on');
AssertEquals_BOOL(Expected := FALSE, Actual := fb_1.OpOut1, Message := 'other outputs off');
AssertEquals_BYTE(Expected := TO_BYTE(E_SafeFbState.Run), Actual := fb_1.State, Message := 'state RUN');
// act: second input also set
group_1(Run := TRUE);
fb_1(OpIn1 := TRUE, OpIn2 := TRUE);
AssertEquals_BOOL(Expected := FALSE, Actual := fb_1.OpOut2, Message := 'all outputs off with two modes selected');
AssertEquals_BYTE(Expected := TO_BYTE(E_SafeFbState.Safe), Actual := fb_1.State, Message := 'state SAFE');
TEST_FINISHED_NAMED(__POUNAME());
END_METHOD

METHOD PRIVATE Test_SlowModeChangeGivesDiscrepancyError
TcUnit.TEST(__POUNAME());
waitTimer_3();

CASE state_3 OF
    10:
        // arrange: mode 1 selected and running
        group_3(Run := TRUE);
        fb_3(OpIn1 := TRUE, OpIn2 := FALSE);
        group_3(Run := TRUE);
        fb_3(OpIn1 := TRUE, OpIn2 := FALSE);
        state_3 := 20;
        waitTimer_3(IN := TRUE, PT := T#250MS);
    20:
        // act: leave mode 1 without selecting another
        group_3(Run := TRUE);
        fb_3(OpIn1 := FALSE, OpIn2 := FALSE);

        IF NOT waitTimer_3.Q THEN
            RETURN;
        END_IF

        waitTimer_3(IN := FALSE);
        // assert
        AssertEquals_BOOL(Expected := TRUE, Actual := fb_3.Error, Message := 'discrepancy error after time without a mode');
        AssertEquals_BYTE(Expected := TO_BYTE(E_SafeFbState.Error), Actual := fb_3.State, Message := 'state ERROR');
        AssertEquals_WORD(Expected := WORD#1, Actual := fb_3.Diag, Message := 'diag bit 0');
        TEST_FINISHED_NAMED(__POUNAME());
        state_3 := 10;
END_CASE
END_METHOD

METHOD PRIVATE Test_OneConnectedInputIsRefused
TcUnit.TEST(__POUNAME());
// arrange / act: OpIn1 is the only connected input, which the Safety Editor refuses
group_4(Run := TRUE);
fb_4(OpIn1 := TRUE);
group_4(Run := TRUE);
fb_4(OpIn1 := TRUE);
// assert
AssertEquals_BOOL(Expected := TRUE, Actual := fb_4.Error, Message := 'configuration error reported');
AssertEquals_BYTE(Expected := TO_BYTE(E_SafeFbState.Error), Actual := fb_4.State, Message := 'state ERROR');
AssertEquals_WORD(Expected := WORD#16#8000, Actual := fb_4.Diag, Message := 'diag bit 15 configuration refused');
AssertEquals_BOOL(Expected := FALSE, Actual := fb_4.OpOut1, Message := 'OpOut1 stays at its safe value');
AssertEquals_BOOL(Expected := TRUE, Actual := group_4.FbErr, Message := 'the group sees an FB error');
// act: ErrAck 0 -> 1 -> 0 does not clear a configuration error
group_4(Run := TRUE, ErrAck := TRUE);
fb_4(OpIn1 := TRUE);
group_4(Run := TRUE, ErrAck := TRUE);
fb_4(OpIn1 := TRUE);
group_4(Run := TRUE, ErrAck := FALSE);
fb_4(OpIn1 := TRUE);
AssertEquals_BOOL(Expected := TRUE, Actual := fb_4.Error, Message := 'error not acknowledged');
AssertEquals_WORD(Expected := WORD#16#8000, Actual := fb_4.Diag, Message := 'diag bit 15 kept');
TEST_FINISHED_NAMED(__POUNAME());
END_METHOD

END_FUNCTION_BLOCK

// ---- FunctionBlocks/T_SafeOpMode.TcPOU
// Model of the TwinSAFE FB OPMODE (operating mode selector).
// Exactly one connected OpIn input must be TRUE for the matching OpOut to be set.
// Manual restart is active when the Restart port is connected.
// The Safety Editor refuses an OPMODE with fewer than two OpIn ports connected: the model then reports
// Error with diagnostic bit 15 instead of running (see T_SafeFunctionBlockBase).
{attribute 'reflection'}
FUNCTION_BLOCK T_SafeOpMode EXTENDS T_SafeFunctionBlockBase
VAR_INPUT
    Restart : BOOL; // may be a standard PLC signal
    OpIn1 : BOOL;
    OpIn2 : BOOL;
    OpIn3 : BOOL;
    OpIn4 : BOOL;
    OpIn5 : BOOL;
    OpIn6 : BOOL;
    OpIn7 : BOOL;
    OpIn8 : BOOL;
    Parameters : ST_SafeOpModeParameters;
END_VAR
VAR_OUTPUT
    OpOut1 : BOOL;
    OpOut2 : BOOL;
    OpOut3 : BOOL;
    OpOut4 : BOOL;
    OpOut5 : BOOL;
    OpOut6 : BOOL;
    OpOut7 : BOOL;
    OpOut8 : BOOL;
END_VAR
VAR
    {attribute 'is_connected' := 'Restart'}
    _restartConnected : BOOL;
    {attribute 'is_connected' := 'OpIn1'}
    _opIn1Connected : BOOL;
    {attribute 'is_connected' := 'OpIn2'}
    _opIn2Connected : BOOL;
    {attribute 'is_connected' := 'OpIn3'}
    _opIn3Connected : BOOL;
    {attribute 'is_connected' := 'OpIn4'}
    _opIn4Connected : BOOL;
    {attribute 'is_connected' := 'OpIn5'}
    _opIn5Connected : BOOL;
    {attribute 'is_connected' := 'OpIn6'}
    _opIn6Connected : BOOL;
    {attribute 'is_connected' := 'OpIn7'}
    _opIn7Connected : BOOL;
    {attribute 'is_connected' := 'OpIn8'}
    _opIn8Connected : BOOL;
    _state : E_SafeFbState := E_SafeFbState.Stop;
    _prevState : E_SafeFbState;
    _restartPrev : BOOL;
    _discrepancyTimer : TON;
    _modeSelectedBefore : BOOL;
END_VAR

SUPER^();

// At least two OpIn ports must be connected (Safety Editor: "OPMODE does not have at least 2 input ports connected").
METHOD PROTECTED ConfigurationOk : BOOL
VAR
    connectedInputs : USINT;
END_VAR
connectedInputs := BOOL_TO_USINT(_opIn1Connected)
    + BOOL_TO_USINT(_opIn2Connected)
    + BOOL_TO_USINT(_opIn3Connected)
    + BOOL_TO_USINT(_opIn4Connected)
    + BOOL_TO_USINT(_opIn5Connected)
    + BOOL_TO_USINT(_opIn6Connected)
    + BOOL_TO_USINT(_opIn7Connected)
    + BOOL_TO_USINT(_opIn8Connected);

IF connectedInputs < 2 THEN
    _configurationFault := 'T_SafeOpMode: OPMODE does not have at least 2 input ports connected';
    RETURN;
END_IF

ConfigurationOk := TRUE;
END_METHOD

METHOD PROTECTED Process
VAR
    count : USINT;
    selected : USINT;
    exactlyOne : BOOL;
    restartFalling : BOOL;
    monitoring : BOOL;
    operating : BOOL;
    stateBefore : E_SafeFbState;
    passes : USINT;
END_VAR
IF _opIn1Connected AND OpIn1 THEN
    count    := count + 1;
    selected := 1;
END_IF

IF _opIn2Connected AND OpIn2 THEN
    count    := count + 1;
    selected := 2;
END_IF

IF _opIn3Connected AND OpIn3 THEN
    count    := count + 1;
    selected := 3;
END_IF

IF _opIn4Connected AND OpIn4 THEN
    count    := count + 1;
    selected := 4;
END_IF

IF _opIn5Connected AND OpIn5 THEN
    count    := count + 1;
    selected := 5;
END_IF

IF _opIn6Connected AND OpIn6 THEN
    count    := count + 1;
    selected := 6;
END_IF

IF _opIn7Connected AND OpIn7 THEN
    count    := count + 1;
    selected := 7;
END_IF

IF _opIn8Connected AND OpIn8 THEN
    count    := count + 1;
    selected := 8;
END_IF

exactlyOne     := (count = 1);
restartFalling := NOT Restart AND _restartPrev;
_restartPrev   := Restart;

IF NOT _fbRun AND _state <> E_SafeFbState.Error AND _state <> E_SafeFbState.Reset THEN
    _state := E_SafeFbState.Stop;
END_IF

// Discrepancy monitoring of a mode change: none or several inputs set for too long
operating  := (_state = E_SafeFbState.Safe) OR (_state = E_SafeFbState.Start) OR (_state = E_SafeFbState.Run);
monitoring := operating AND _modeSelectedBefore AND NOT exactlyOne AND (Parameters.DiscrepancyTime > T#0S);
_discrepancyTimer(IN := monitoring, PT := Parameters.DiscrepancyTime);

IF _discrepancyTimer.Q AND operating THEN
    SetDiagBit(0);
    _state := E_SafeFbState.Error;
END_IF

passes := 0;

REPEAT
    stateBefore := _state;

    CASE _state OF
        E_SafeFbState.Stop:
            IF StateChanged() THEN
                SetOutputs(0);
                Error               := FALSE;
                Diag                := 0;
                _modeSelectedBefore := FALSE;
            END_IF

            IF _fbRun THEN
                _state := E_SafeFbState.Safe;
            END_IF

        E_SafeFbState.Safe:
            IF StateChanged() THEN
                SetOutputs(0);
            END_IF

            IF exactlyOne THEN
                IF NOT _restartConnected THEN
                    _state := E_SafeFbState.Run;
                ELSIF Restart THEN
                    _state := E_SafeFbState.Start;
                END_IF
            END_IF

        E_SafeFbState.Start:
            IF StateChanged() THEN
                SetOutputs(0);
            END_IF

            IF NOT exactlyOne THEN
                _state := E_SafeFbState.Safe;
            ELSIF restartFalling THEN
                _state := E_SafeFbState.Run;
            END_IF

        E_SafeFbState.Run:
            IF StateChanged() THEN
                _modeSelectedBefore := TRUE;
            END_IF

            IF exactlyOne THEN
                SetOutputs(selected);
            ELSE
                SetOutputs(0);
                _state := E_SafeFbState.Safe;
            END_IF

        E_SafeFbState.Error:
            IF StateChanged() THEN
                SetOutputs(0);
                Error := TRUE;
            END_IF

            IF _errAck THEN
                _state := E_SafeFbState.Reset;
            END_IF

        E_SafeFbState.Reset:
            IF StateChanged() THEN
                Error := FALSE;
                Diag  := 0;
            END_IF

            IF _errAckFallingEdge THEN
                _state := SEL(_fbRun, E_SafeFbState.Stop, E_SafeFbState.Safe);
            END_IF
    END_CASE

    passes := passes + 1;
UNTIL (stateBefore = _state) OR (passes >= 3)
END_REPEAT

State := TO_BYTE(_state);
END_METHOD

METHOD PRIVATE SetOutputs
VAR_INPUT
    selected : USINT; // 0 = all outputs off
END_VAR
OpOut1 := (selected = 1);
OpOut2 := (selected = 2);
OpOut3 := (selected = 3);
OpOut4 := (selected = 4);
OpOut5 := (selected = 5);
OpOut6 := (selected = 6);
OpOut7 := (selected = 7);
OpOut8 := (selected = 8);
END_METHOD

METHOD PRIVATE StateChanged : BOOL
IF _prevState = _state THEN
    RETURN;
END_IF

_prevState   := _state;
StateChanged := TRUE;
END_METHOD

END_FUNCTION_BLOCK

// ---- Tests/T_SafeRs_Tests.TcPOU
FUNCTION_BLOCK T_SafeRs_Tests EXTENDS TcUnit.FB_TestSuite
VAR
    // Test_ResetDominantLatch
    group_1 : T_SafeGroup;
    fb_1 : T_SafeRs(group := group_1);
    // Test_UnconnectedSetIsRefused
    group_2 : T_SafeGroup;
    fb_2 : T_SafeRs(group := group_2);
END_VAR

Test_ResetDominantLatch();
Test_UnconnectedSetIsRefused();

METHOD PRIVATE Test_ResetDominantLatch
TcUnit.TEST(__POUNAME());
// act / assert
group_1(Run := TRUE);
fb_1(Set := TRUE, Reset := FALSE);
AssertEquals_BOOL(Expected := TRUE, Actual := fb_1.RsOut, Message := 'set');
fb_1(Set := FALSE, Reset := FALSE);
AssertEquals_BOOL(Expected := TRUE, Actual := fb_1.RsOut, Message := 'held');
fb_1(Set := TRUE, Reset := TRUE);
AssertEquals_BOOL(Expected := FALSE, Actual := fb_1.RsOut, Message := 'reset dominant');
TEST_FINISHED_NAMED(__POUNAME());
END_METHOD

METHOD PRIVATE Test_UnconnectedSetIsRefused
TcUnit.TEST(__POUNAME());
// arrange / act: Set is unconnected, which the Safety Editor refuses
group_2(Run := TRUE);
fb_2(Reset := FALSE);
group_2(Run := TRUE);
fb_2(Reset := FALSE);
// assert
AssertEquals_BOOL(Expected := TRUE, Actual := fb_2.Error, Message := 'configuration error reported');
AssertEquals_BYTE(Expected := TO_BYTE(E_SafeFbState.Error), Actual := fb_2.State, Message := 'state ERROR');
AssertEquals_WORD(Expected := WORD#16#8000, Actual := fb_2.Diag, Message := 'diag bit 15 configuration refused');
AssertEquals_BOOL(Expected := FALSE, Actual := fb_2.RsOut, Message := 'RsOut stays at its safe value');
AssertEquals_BOOL(Expected := TRUE, Actual := group_2.FbErr, Message := 'the group sees an FB error');
// act: ErrAck 0 -> 1 -> 0 does not clear a configuration error
group_2(Run := TRUE, ErrAck := TRUE);
fb_2(Reset := FALSE);
group_2(Run := TRUE, ErrAck := TRUE);
fb_2(Reset := FALSE);
group_2(Run := TRUE, ErrAck := FALSE);
fb_2(Reset := FALSE);
AssertEquals_BOOL(Expected := TRUE, Actual := fb_2.Error, Message := 'error not acknowledged');
AssertEquals_WORD(Expected := WORD#16#8000, Actual := fb_2.Diag, Message := 'diag bit 15 kept');
TEST_FINISHED_NAMED(__POUNAME());
END_METHOD

END_FUNCTION_BLOCK

// ---- FunctionBlocks/T_SafeRs.TcPOU
// Model of the TwinSAFE FB RS (reset dominant latch).
// The Safety Editor refuses an RS with Set or Reset unconnected: the model then reports Error with
// diagnostic bit 15 instead of running (see T_SafeFunctionBlockBase).
{attribute 'reflection'}
FUNCTION_BLOCK T_SafeRs EXTENDS T_SafeFunctionBlockBase
VAR_INPUT
    Set : BOOL;
    Reset : BOOL;
    Parameters : ST_SafeLatchParameters;
END_VAR
VAR_OUTPUT
    RsOut : BOOL;
END_VAR
VAR
    {attribute 'is_connected' := 'Set'}
    _setConnected : BOOL;
    {attribute 'is_connected' := 'Reset'}
    _resetConnected : BOOL;
    _state : E_SafeLatchState := E_SafeLatchState.Stop;
END_VAR

SUPER^();

// Set and Reset must both be connected (Safety Editor: "Inport Set of RS must be connected").
METHOD PROTECTED ConfigurationOk : BOOL
IF NOT _setConnected THEN
    _configurationFault := 'T_SafeRs: Inport Set of RS must be connected';
    RETURN;
ELSIF NOT _resetConnected THEN
    _configurationFault := 'T_SafeRs: Inport Reset of RS must be connected';
    RETURN;
END_IF

ConfigurationOk := TRUE;
END_METHOD

METHOD PROTECTED Process
VAR
    setActive : BOOL;
    resetActive : BOOL;
END_VAR
setActive   := F_SafeInputValue(_setConnected, Parameters.SetMakeContact, Set);
resetActive := F_SafeInputValue(_resetConnected, Parameters.ResetMakeContact, Reset);

IF NOT _fbRun THEN
    _state := E_SafeLatchState.Stop;
ELSE
    IF _state = E_SafeLatchState.Stop THEN
        _state := E_SafeLatchState.Safe;
    END_IF

    IF resetActive THEN
        _state := E_SafeLatchState.Safe;
    ELSIF setActive THEN
        _state := E_SafeLatchState.Set;
    END_IF
END_IF

RsOut := (_state = E_SafeLatchState.Set);
Error := FALSE;
Diag  := 0;
State := TO_BYTE(_state);
END_METHOD

END_FUNCTION_BLOCK

// ---- Tests/T_SafeSr_Tests.TcPOU
FUNCTION_BLOCK T_SafeSr_Tests EXTENDS TcUnit.FB_TestSuite
VAR
    // Test_SetDominantLatch
    group_1 : T_SafeGroup;
    fb_1 : T_SafeSr(group := group_1);
    // Test_UnconnectedResetIsRefused
    group_2 : T_SafeGroup;
    fb_2 : T_SafeSr(group := group_2);
END_VAR

Test_SetDominantLatch();
Test_UnconnectedResetIsRefused();

METHOD PRIVATE Test_SetDominantLatch
TcUnit.TEST(__POUNAME());
// act / assert
group_1(Run := TRUE);
fb_1(Set := TRUE, Reset := TRUE);
AssertEquals_BOOL(Expected := TRUE, Actual := fb_1.SrOut, Message := 'set dominant');
fb_1(Set := FALSE, Reset := TRUE);
AssertEquals_BOOL(Expected := FALSE, Actual := fb_1.SrOut, Message := 'reset');
fb_1(Set := FALSE, Reset := FALSE);
AssertEquals_BOOL(Expected := FALSE, Actual := fb_1.SrOut, Message := 'held');
TEST_FINISHED_NAMED(__POUNAME());
END_METHOD

METHOD PRIVATE Test_UnconnectedResetIsRefused
TcUnit.TEST(__POUNAME());
// arrange / act: Reset is unconnected, which the Safety Editor refuses
group_2(Run := TRUE);
fb_2(Set := TRUE);
group_2(Run := TRUE);
fb_2(Set := TRUE);
// assert
AssertEquals_BOOL(Expected := TRUE, Actual := fb_2.Error, Message := 'configuration error reported');
AssertEquals_BYTE(Expected := TO_BYTE(E_SafeFbState.Error), Actual := fb_2.State, Message := 'state ERROR');
AssertEquals_WORD(Expected := WORD#16#8000, Actual := fb_2.Diag, Message := 'diag bit 15 configuration refused');
AssertEquals_BOOL(Expected := FALSE, Actual := fb_2.SrOut, Message := 'SrOut stays at its safe value');
AssertEquals_BOOL(Expected := TRUE, Actual := group_2.FbErr, Message := 'the group sees an FB error');
// act: ErrAck 0 -> 1 -> 0 does not clear a configuration error
group_2(Run := TRUE, ErrAck := TRUE);
fb_2(Set := TRUE);
group_2(Run := TRUE, ErrAck := TRUE);
fb_2(Set := TRUE);
group_2(Run := TRUE, ErrAck := FALSE);
fb_2(Set := TRUE);
AssertEquals_BOOL(Expected := TRUE, Actual := fb_2.Error, Message := 'error not acknowledged');
AssertEquals_WORD(Expected := WORD#16#8000, Actual := fb_2.Diag, Message := 'diag bit 15 kept');
TEST_FINISHED_NAMED(__POUNAME());
END_METHOD

END_FUNCTION_BLOCK

// ---- FunctionBlocks/T_SafeSr.TcPOU
// Model of the TwinSAFE FB SR (set dominant latch).
// The Safety Editor refuses an SR with Set or Reset unconnected: the model then reports Error with
// diagnostic bit 15 instead of running (see T_SafeFunctionBlockBase).
{attribute 'reflection'}
FUNCTION_BLOCK T_SafeSr EXTENDS T_SafeFunctionBlockBase
VAR_INPUT
    Set : BOOL;
    Reset : BOOL;
    Parameters : ST_SafeLatchParameters;
END_VAR
VAR_OUTPUT
    SrOut : BOOL;
END_VAR
VAR
    {attribute 'is_connected' := 'Set'}
    _setConnected : BOOL;
    {attribute 'is_connected' := 'Reset'}
    _resetConnected : BOOL;
    _state : E_SafeLatchState := E_SafeLatchState.Stop;
END_VAR

SUPER^();

// Set and Reset must both be connected (Safety Editor: "Inport Set of SR must be connected").
METHOD PROTECTED ConfigurationOk : BOOL
IF NOT _setConnected THEN
    _configurationFault := 'T_SafeSr: Inport Set of SR must be connected';
    RETURN;
ELSIF NOT _resetConnected THEN
    _configurationFault := 'T_SafeSr: Inport Reset of SR must be connected';
    RETURN;
END_IF

ConfigurationOk := TRUE;
END_METHOD

METHOD PROTECTED Process
VAR
    setActive : BOOL;
    resetActive : BOOL;
END_VAR
setActive   := F_SafeInputValue(_setConnected, Parameters.SetMakeContact, Set);
resetActive := F_SafeInputValue(_resetConnected, Parameters.ResetMakeContact, Reset);

IF NOT _fbRun THEN
    _state := E_SafeLatchState.Stop;
ELSE
    IF _state = E_SafeLatchState.Stop THEN
        _state := E_SafeLatchState.Safe;
    END_IF

    IF setActive THEN
        _state := E_SafeLatchState.Set;
    ELSIF resetActive THEN
        _state := E_SafeLatchState.Safe;
    END_IF
END_IF

SrOut := (_state = E_SafeLatchState.Set);
Error := FALSE;
Diag  := 0;
State := TO_BYTE(_state);
END_METHOD

END_FUNCTION_BLOCK

// ---- Tests/T_SafeTon_Tests.TcPOU
FUNCTION_BLOCK T_SafeTon_Tests EXTENDS TcUnit.FB_TestSuite
VAR
    // Test_OutputDelayedOn
    group_1 : T_SafeGroup;
    fb_1 : T_SafeTon(group := group_1) := (Parameters := (DelayTime := T#100MS));
    state_1 : INT := 10;
    waitTimer_1 : TON;
    // Test_UnconnectedInputIsRefused
    group_2 : T_SafeGroup;
    fb_2 : T_SafeTon(group := group_2);
END_VAR

Test_OutputDelayedOn();
Test_UnconnectedInputIsRefused();

METHOD PRIVATE Test_OutputDelayedOn
TcUnit.TEST(__POUNAME());
waitTimer_1();

CASE state_1 OF
    10:
        // act
        group_1(Run := TRUE);
        fb_1(TonIn1 := TRUE);
        // assert
        AssertEquals_BOOL(Expected := FALSE, Actual := fb_1.TonOut, Message := 'output not yet on');
        AssertEquals_BYTE(Expected := TO_BYTE(E_SafeTonState.DelayIn), Actual := fb_1.State, Message := 'state DELAYIN');
        state_1 := 20;
        waitTimer_1(IN := TRUE, PT := T#200MS);
    20:
        group_1(Run := TRUE);
        fb_1(TonIn1 := TRUE);

        IF NOT waitTimer_1.Q THEN
            RETURN;
        END_IF

        waitTimer_1(IN := FALSE);
        // assert
        AssertEquals_BOOL(Expected := TRUE, Actual := fb_1.TonOut, Message := 'output on after the delay');
        fb_1(TonIn1 := FALSE);
        AssertEquals_BOOL(Expected := FALSE, Actual := fb_1.TonOut, Message := 'output off immediately');
        TEST_FINISHED_NAMED(__POUNAME());
        state_1 := 10;
END_CASE
END_METHOD

METHOD PRIVATE Test_UnconnectedInputIsRefused
TcUnit.TEST(__POUNAME());
// arrange / act: TonIn1 is unconnected, which the Safety Editor refuses
group_2(Run := TRUE);
fb_2();
group_2(Run := TRUE);
fb_2();
// assert
AssertEquals_BOOL(Expected := TRUE, Actual := fb_2.Error, Message := 'configuration error reported');
AssertEquals_BYTE(Expected := TO_BYTE(E_SafeFbState.Error), Actual := fb_2.State, Message := 'state ERROR');
AssertEquals_WORD(Expected := WORD#16#8000, Actual := fb_2.Diag, Message := 'diag bit 15 configuration refused');
AssertEquals_BOOL(Expected := FALSE, Actual := fb_2.TonOut, Message := 'TonOut stays at its safe value');
AssertEquals_BOOL(Expected := TRUE, Actual := group_2.FbErr, Message := 'the group sees an FB error');
// act: ErrAck 0 -> 1 -> 0 does not clear a configuration error
group_2(Run := TRUE, ErrAck := TRUE);
fb_2();
group_2(Run := TRUE, ErrAck := TRUE);
fb_2();
group_2(Run := TRUE, ErrAck := FALSE);
fb_2();
AssertEquals_BOOL(Expected := TRUE, Actual := fb_2.Error, Message := 'error not acknowledged');
AssertEquals_WORD(Expected := WORD#16#8000, Actual := fb_2.Diag, Message := 'diag bit 15 kept');
TEST_FINISHED_NAMED(__POUNAME());
END_METHOD

END_FUNCTION_BLOCK

// ---- FunctionBlocks/T_SafeTon.TcPOU
// Model of the TwinSAFE FB TON (switch-on delay).
// The Safety Editor refuses a TON with TonIn1 unconnected: the model then reports Error with diagnostic
// bit 15 instead of running (see T_SafeFunctionBlockBase).
{attribute 'reflection'}
FUNCTION_BLOCK T_SafeTon EXTENDS T_SafeFunctionBlockBase
VAR_INPUT
    TonIn1 : BOOL;
    Parameters : ST_SafeTimerParameters;
END_VAR
VAR_OUTPUT
    TonOut : BOOL;
END_VAR
VAR
    {attribute 'is_connected' := 'TonIn1'}
    _tonIn1Connected : BOOL;
    _state : E_SafeTonState := E_SafeTonState.Stop;
    _timer : TON;
END_VAR

SUPER^();

// TonIn1 must be connected (Safety Editor: "Inport TonIn1 of TON must be connected").
METHOD PROTECTED ConfigurationOk : BOOL
IF NOT _tonIn1Connected THEN
    _configurationFault := 'T_SafeTon: Inport TonIn1 of TON must be connected';
    RETURN;
END_IF

ConfigurationOk := TRUE;
END_METHOD

METHOD PROTECTED Process
VAR
    inputActive : BOOL;
END_VAR
inputActive := _fbRun AND F_SafeInputValue(_tonIn1Connected, Parameters.MakeContact, TonIn1);
_timer(IN := inputActive, PT := Parameters.DelayTime);

IF NOT _fbRun THEN
    _state := E_SafeTonState.Stop;
ELSIF NOT inputActive THEN
    _state := E_SafeTonState.Safe;
ELSIF _timer.Q THEN
    _state := E_SafeTonState.Run;
ELSE
    _state := E_SafeTonState.DelayIn;
END_IF

TonOut := (_state = E_SafeTonState.Run);
Error  := FALSE;
Diag   := 0;
State  := TO_BYTE(_state);
END_METHOD

END_FUNCTION_BLOCK

// ---- Tests/T_SafeTof_Tests.TcPOU
FUNCTION_BLOCK T_SafeTof_Tests EXTENDS TcUnit.FB_TestSuite
VAR
    // Test_OutputDelayedOff
    group_1 : T_SafeGroup;
    fb_1 : T_SafeTof(group := group_1) := (Parameters := (DelayTime := T#100MS));
    state_1 : INT := 10;
    waitTimer_1 : TON;
    // Test_UnconnectedInputIsRefused
    group_2 : T_SafeGroup;
    fb_2 : T_SafeTof(group := group_2);
END_VAR

Test_OutputDelayedOff();
Test_UnconnectedInputIsRefused();

METHOD PRIVATE Test_OutputDelayedOff
TcUnit.TEST(__POUNAME());
waitTimer_1();

CASE state_1 OF
    10:
        group_1(Run := TRUE);
        fb_1(TofIn1 := TRUE);
        AssertEquals_BOOL(Expected := TRUE, Actual := fb_1.TofOut, Message := 'output on immediately');
        // act
        fb_1(TofIn1 := FALSE);
        AssertEquals_BOOL(Expected := TRUE, Actual := fb_1.TofOut, Message := 'output held during the delay');
        AssertEquals_BYTE(Expected := TO_BYTE(E_SafeFbState.DelayOut), Actual := fb_1.State, Message := 'state DELAYOUT');
        state_1 := 20;
        waitTimer_1(IN := TRUE, PT := T#200MS);
    20:
        group_1(Run := TRUE);
        fb_1(TofIn1 := FALSE);

        IF NOT waitTimer_1.Q THEN
            RETURN;
        END_IF

        waitTimer_1(IN := FALSE);
        // assert
        AssertEquals_BOOL(Expected := FALSE, Actual := fb_1.TofOut, Message := 'output off after the delay');
        TEST_FINISHED_NAMED(__POUNAME());
        state_1 := 10;
END_CASE
END_METHOD

METHOD PRIVATE Test_UnconnectedInputIsRefused
TcUnit.TEST(__POUNAME());
// arrange / act: TofIn1 is unconnected, which the Safety Editor refuses
group_2(Run := TRUE);
fb_2();
group_2(Run := TRUE);
fb_2();
// assert
AssertEquals_BOOL(Expected := TRUE, Actual := fb_2.Error, Message := 'configuration error reported');
AssertEquals_BYTE(Expected := TO_BYTE(E_SafeFbState.Error), Actual := fb_2.State, Message := 'state ERROR');
AssertEquals_WORD(Expected := WORD#16#8000, Actual := fb_2.Diag, Message := 'diag bit 15 configuration refused');
AssertEquals_BOOL(Expected := FALSE, Actual := fb_2.TofOut, Message := 'TofOut stays at its safe value');
AssertEquals_BOOL(Expected := TRUE, Actual := group_2.FbErr, Message := 'the group sees an FB error');
// act: ErrAck 0 -> 1 -> 0 does not clear a configuration error
group_2(Run := TRUE, ErrAck := TRUE);
fb_2();
group_2(Run := TRUE, ErrAck := TRUE);
fb_2();
group_2(Run := TRUE, ErrAck := FALSE);
fb_2();
AssertEquals_BOOL(Expected := TRUE, Actual := fb_2.Error, Message := 'error not acknowledged');
AssertEquals_WORD(Expected := WORD#16#8000, Actual := fb_2.Diag, Message := 'diag bit 15 kept');
TEST_FINISHED_NAMED(__POUNAME());
END_METHOD

END_FUNCTION_BLOCK

// ---- FunctionBlocks/T_SafeTof.TcPOU
// Model of the TwinSAFE FB TOF (switch-off delay).
// The Safety Editor refuses a TOF with TofIn1 unconnected: the model then reports Error with diagnostic
// bit 15 instead of running (see T_SafeFunctionBlockBase).
{attribute 'reflection'}
FUNCTION_BLOCK T_SafeTof EXTENDS T_SafeFunctionBlockBase
VAR_INPUT
    TofIn1 : BOOL;
    Parameters : ST_SafeTimerParameters;
END_VAR
VAR_OUTPUT
    TofOut : BOOL;
END_VAR
VAR
    {attribute 'is_connected' := 'TofIn1'}
    _tofIn1Connected : BOOL;
    _state : E_SafeFbState := E_SafeFbState.Stop;
    _timer : TOF;
END_VAR

SUPER^();

// TofIn1 must be connected (Safety Editor: "Inport TofIn1 of TOF must be connected").
METHOD PROTECTED ConfigurationOk : BOOL
IF NOT _tofIn1Connected THEN
    _configurationFault := 'T_SafeTof: Inport TofIn1 of TOF must be connected';
    RETURN;
END_IF

ConfigurationOk := TRUE;
END_METHOD

METHOD PROTECTED Process
VAR
    inputActive : BOOL;
END_VAR
inputActive := F_SafeInputValue(_tofIn1Connected, Parameters.MakeContact, TofIn1);

IF NOT _fbRun THEN
    // a stopped FB does not run its delay
    _timer(IN := FALSE, PT := T#0S);
    _state := E_SafeFbState.Stop;
ELSE
    _timer(IN := inputActive, PT := Parameters.DelayTime);

    IF inputActive THEN
        _state := E_SafeFbState.Run;
    ELSIF _timer.Q THEN
        _state := E_SafeFbState.DelayOut;
    ELSE
        _state := E_SafeFbState.Safe;
    END_IF
END_IF

TofOut := (_state = E_SafeFbState.Run) OR (_state = E_SafeFbState.DelayOut);
Error  := FALSE;
Diag   := 0;
State  := TO_BYTE(_state);
END_METHOD

END_FUNCTION_BLOCK

// ---- Tests/T_SafeEdm_Tests.TcPOU
FUNCTION_BLOCK T_SafeEdm_Tests EXTENDS TcUnit.FB_TestSuite
VAR
    // Test_SwitchOnTimeoutGivesError
    group_1 : T_SafeGroup;
    fb_1 : T_SafeEdm(group := group_1) := (Parameters := (SwitchOnTime := T#100MS));
    state_1 : INT := 10;
    waitTimer_1 : TON;
    // Test_NoErrorWhenFeedbackFollows
    group_2 : T_SafeGroup;
    fb_2 : T_SafeEdm(group := group_2) := (Parameters := (SwitchOnTime := T#100MS, SwitchOffTime := T#100MS));
    state_2 : INT := 10;
    waitTimer_2 : TON;
    // Test_UnconnectedMon2IsRefused
    group_3 : T_SafeGroup;
    fb_3 : T_SafeEdm(group := group_3);
END_VAR

Test_SwitchOnTimeoutGivesError();
Test_NoErrorWhenFeedbackFollows();
Test_UnconnectedMon2IsRefused();

METHOD PRIVATE Test_NoErrorWhenFeedbackFollows
TcUnit.TEST(__POUNAME());
waitTimer_2();

CASE state_2 OF
    10:
        state_2 := 20;
        waitTimer_2(IN := TRUE, PT := T#200MS);
    20:
        group_2(Run := TRUE);
        fb_2(Mon1 := TRUE, Mon2 := FALSE);

        IF NOT waitTimer_2.Q THEN
            RETURN;
        END_IF

        waitTimer_2(IN := FALSE);
        AssertEquals_BOOL(Expected := FALSE, Actual := fb_2.Error, Message := 'no error while feedback is correct');
        state_2 := 30;
        waitTimer_2(IN := TRUE, PT := T#200MS);
    30:
        // act: switch off, feedback follows immediately
        group_2(Run := TRUE);
        fb_2(Mon1 := FALSE, Mon2 := TRUE);

        IF NOT waitTimer_2.Q THEN
            RETURN;
        END_IF

        waitTimer_2(IN := FALSE);
        AssertEquals_BOOL(Expected := FALSE, Actual := fb_2.Error, Message := 'no error after switch-off with feedback');
        TEST_FINISHED_NAMED(__POUNAME());
        state_2 := 10;
END_CASE
END_METHOD

METHOD PRIVATE Test_SwitchOnTimeoutGivesError
TcUnit.TEST(__POUNAME());
waitTimer_1();

CASE state_1 OF
    10:
        state_1 := 20;
        waitTimer_1(IN := TRUE, PT := T#250MS);
    20:
        // act: Mon1 on, feedback never follows
        group_1(Run := TRUE, ErrAck := FALSE);
        fb_1(Mon1 := TRUE, Mon2 := TRUE);

        IF NOT waitTimer_1.Q THEN
            RETURN;
        END_IF

        waitTimer_1(IN := FALSE);
        // assert
        AssertEquals_BOOL(Expected := TRUE, Actual := fb_1.Error, Message := 'error when Mon2 does not drop in time');
        AssertEquals_WORD(Expected := WORD#2, Actual := fb_1.Diag, Message := 'diag bit 1 switch-on timer elapsed');
        // act: acknowledge (two cycles raised so the group_1 reaches RESET, then released)
        group_1(Run := TRUE, ErrAck := TRUE);
        fb_1(Mon1 := TRUE, Mon2 := TRUE);
        group_1(Run := TRUE, ErrAck := TRUE);
        fb_1(Mon1 := TRUE, Mon2 := TRUE);
        group_1(Run := TRUE, ErrAck := FALSE);
        fb_1(Mon1 := TRUE, Mon2 := FALSE);
        AssertEquals_BOOL(Expected := FALSE, Actual := fb_1.Error, Message := 'error cleared after acknowledgement');
        TEST_FINISHED_NAMED(__POUNAME());
        state_1 := 10;
END_CASE
END_METHOD

